	fbController				:FB_STOEBER_AxisController;
	fbMoveManual				:FB_STOEBER_AxisMoveManual;
	fbMoveAuto					:FB_STOEBER_AxisMoveAuto;
	(*fbDriveLink				:FB_STOEBER_DriveLink;*)
	fbForce						:FB_ScalingOffset;
	fbForceCtrl					:FB_ForceController;
	fbCoolingOff				:FB_SignalHandlingDelay;
	
	fbSawingOverride			:FB_Override;
	rtWriteForcePara			:R_TRIG;
	
	fbForceSimple				:FB_ScalingOffset;
	fbForceEL3351				:FB_EL3351;
	fbForceEL3356				:FB_EL3356;

	
END_VAR


IF NOT bEnable								(* Signal FB enable *)
THEN
	bCtrlEnabled := TRUE;
	bReferenced := TRUE;
	bNotMoving := TRUE;
	
	RETURN;
END_IF

A_AxisLink();
A_AxisGetStatus();
A_AxisController();
A_AxisForceCtrl();
A_AxisMoveManual();
A_AxisMoveAuto();
A_AxisTerminalDiag();
A_AxisAlarm();

ACTION A_AxisAlarm:

(* Axis error *)
tonAxisEnabled(
	IN := fbController.bEnable
		AND fbController.bRegulatorOn
		AND NOT fbController.bStatusDelay,
	PT := fbController.tStatusDelay + t#2s
);

bErrorCtrlEnabled := tonAxisEnabled.Q;
(*byErrorPLCOpenController := fbAxisControl.byPLCOpenErrCode;*)
(*bErrorController := fbAxisControl.bError;
bErrorMoveManual := fbMoveManual.bError;
bErrorMoveAuto := fbMoveAuto.bError;*)
END_ACTION

ACTION A_AxisController:

(* Axis controller *)
fbController(
    bEnable := TRUE,
	etMachineMode := etMachineMode,
	etMachineState := etMachineState,
	bNoEStop := bNoEStop,
	bRegulatorOn := bNoEStop
				      AND bPowerSupplyOn
				      AND bSafetyOk
				      AND SEL(bNotMoving, NOT bCtrlInterrupt, TRUE)
				      AND NOT fbMoveManual.bControllerOff
				      AND NOT fbMoveAuto.bControllerOff,
	bReset := bConfirmAlarm,
	bTerminalOK := fbTerminalDiagnosis.bTerminalOK,
	bExeReset := bExeReset,
	bExeSetPos := bExeSetPos,
	lrSetPosition := lrTargetPosition,
	bExeGearIn := bExeGearIn,
	bExeGearOut := bExeGearOut,
	dnRatioNumerator := dnRatioNumerator,
	udnRatioDenominator := udnRatioDenominator,
	lrOverride := SEL(bExtOverrideEn,
					SEL(
						bVeloForceCtrlEn,
						lrOverride,
						fbForceCtrl.lrCVVelo),
					lrOverride*lrExtOverride/100.0)/2,
	bWithAbsoluteEncoder := bWithAbsoluteEncoder,
	bPosLagMonitoringEn := bPosLagMonitoringEn,
	lrPositionBias := lrOriginShiftPos,
	lrSoftLimitMax := lrSoftLimitMax,
	lrSoftLimitMin := lrSoftLimitMin,
	bSignalHWLimitMax:= bSignalHWLimitMax,
	bSignalHWLimitMin := bSignalHWLimitMin,
	lrAcceleration := lrAcceleration,
	lrDeceleration := lrDeceleration,
	lrJerk := lrJerk,
	pDrive := ADR(Drive),
	Axis := Axis,
	MasterAxis := MasterAxis,
	bStatusDelay => bCtrlEnabled,
	lrActPos => lrActPosition,
	lrActAbsPos => lrActAbsPosition,
	lrActVelo => lrActVelocity,
	bNotMoving => bNotMoving,
	bStandStill => bStandStill,
	bReferenced => bReferenced,
	bCoupled => bCoupled,
	lrVeloLimitMax => lrVeloMax,
	lrAccLimitMax => lrAccMax,
	lrDecLimitMax => lrDecMax,
	lrJerkLimitMax => lrJerkMax,
	bHardLimitMaxExceeded => bHardLimitMaxExceeded,
	bHardLimitMinExceeded => bHardLimitMinExceeded,
	bSoftLimitMaxExceeded => bSoftLimitMaxExceeded,
	bSoftLimitMinExceeded => bSoftLimitMinExceeded,

);

bSafetyDriveEnable := fbMoveManual.bSafetyCtrlEnable 
				 	  OR fbMoveAuto.bSafetyCtrlEnable;


(* From Tc2)

(* Sawbow sawing override *)
fbSawingOverride(
	bEnable := bExtOverrideEn
			    AND
			    (etgGr00MachineState = ET_MachineState_eAutoExe
			    OR etgGr00MachineState = ET_MachineState_eAutoSteppingExe)
			    AND
			    (etMachineMode = ET_MachineMode_eAutomatic
			     OR etMachineMode = ET_MachineMode_eCycle
			     OR etMachineMode = ET_MachineMode_eStepping),
	bBypassAccDec := FALSE,
	bSetOverideMax := FALSE,
	rSetOverride := rSetSawingOverride,
	rAcc := rgGr00AdsOverrideAcc,
	rDec := rgGr01AdsOverrideDec
);


IF bExtOverrideEn
     AND
    (etgGr00MachineState = ET_MachineState_eAutoExe
    OR etgGr00MachineState = ET_MachineState_eAutoSteppingExe)
    AND
    (etMachineMode = ET_MachineMode_eAutomatic
     OR etMachineMode = ET_MachineMode_eCycle
     OR etMachineMode = ET_MachineMode_eStepping)
THEN
	rSawingOverride := INT_TO_REAL(nSetSawingOverride)/32767.0 * 100.0;
ELSE
	rSawingOverride := 100.0;
END_IF;

(* Axis controller *)
fbController(
    	bEnable := TRUE,
	etMachineMode := etMachineMode,
	etMachineState := etMachineState,
	bRegulatorOn := bNoEStop
				      AND bPowerSupplyOn
				      AND bSafetyOK
                   		      AND NOT bCtrlInterrupt
				      AND NOT fbMoveManual.bControllerOff
				      AND NOT fbMoveAuto.bControllerOff,
	bReset := bConfirmAlarm,
	bCMDInterrupt := bMoveInterrupt,
	bTerminalOK := fbTerminalDiagnosis.bTerminalOK,
	bExeReset := bExeReset,
  	bExeGearIn := bExeGearIn,
    	bExeGearOut := bExeGearOut,
   	dnRatioNumerator := dnRatioNumerator,
    	udnRatioDenominator := udnRatioDenominator,
	lrOverride := SEL(bExtOverrideEn,
					SEL(
						bVeloForceCtrlEn,
						lrOverride,
						fbForceCtrl.lrCVVelo),
					lrOverride * rSawingOverride / 100),
	lrEngineTorque := SEL(
						bEngineTorqueLimitEn,
						nTorqueLimitMax,
						(lrEngineTorque) / 1),
	bWithAbsoluteEncoder := bWithAbsoluteEncoder,
	bHWSignalLimitMax := bHWSignalLimitMax,
	bHWSignalLimitMin := bHWSignalLimitMin,
	lrSoftLimitMax := lrSoftLimitMax,
	lrSoftLimitMin := lrSoftLimitMin,
	lrAcceleration := lrAcceleration,
	lrDeceleration := lrDeceleration,
	lrJerk := lrJerk,
	tTimeOut := tAdsTimeOut,
	Axis := Axis,
	bStatusDelay => bCtrlEnabled,
	lrActPos => lrActPosition,
	lrActVelo => lrActVelocity,
	bNotMoving => bNotMoving,
	bReferenced => bReferenced,
	bCoupled => bCoupled,
	bHardLimitMaxExceeded => bHardLimitMaxExceeded,
	bHardLimitMinExceeded => bHardLimitMinExceeded,
	bSoftLimitMaxExceeded => bSoftLimitMaxExceeded,
	bSoftLimitMinExceeded => bSoftLimitMinExceeded
);

*)
END_ACTION

ACTION A_AxisForceCtrl:

IF unForceMeasureType = 1			(* Current or voltage force measure *)
THEN
	fbForceCtrl.lrMaxForce := lrForceMaxN; (* [N] *)

	fbForceSimple(
		bEnable := TRUE,
		lrInput := lrForceCurrent,
		lrXLowLimit := lrForceMinmA, (* 16#0000 = 4 [mA] *)
		lrXUpperLimit := lrForceMaxmA, (* 16#7FFF = 20 [mA] *)
		lrYLowLimit := lrForceMinN,  (*[N]*)
		lrYUpperLimit := lrForceMaxN,  (*[N]*)
		usiPrecision := 2,
		lrOffset := rForceOffset,
		lrOutputPV => lrActForce
	);


ELSIF unForceMeasureType = 2			(* EL3351 force measure *)
THEN
	fbForceCtrl.lrMaxForce := lrForceMaxN; (* [N] *)

	fbForceEL3351(
		bEnable := TRUE,
		nTerminalNr := 1,
		stTerminalState := ,
		stBridgeState := ,
		stSupplyState := ,
		dnRefvoltage := ,
		dnDiffvoltage := ,
		rOffset := rForceOffset,
		usiPrecision := 2,
		bDeviceOk => ,
		sDeviceStatus => ,
		rUdiff => ,
		rUref => ,
		lrGrossWeightRV=> ,
		lrGrossWeightPV => lrActForce,
		lrNetWeightRV=> ,
		lrNetWeightPV=> ,
		lrTareWeightRV=> ,
		lrTareWeightPV=>
	);

ELSIF  unForceMeasureType = 3			(* EL3356 force measure *)
THEN

(*
	rtWriteForcePara(
		CLK:= bgGr01ForceActiv5kN
			   XOR bgGr01ForceActiv10kN
	);

	CASE nStepWriteForcePara OF
		0:	(*Idle*)

			fbForceEL3356.bWriteCoePara:= FALSE;
			bWriteForceParaBusy := FALSE;

			IF rtWriteForcePara.Q
			THEN
				nStepWriteForcePara := 10;
				bWriteForceParaBusy := TRUE;
			END_IF
		10: 	(*Start*)

			IF bgGr01ForceActiv5kN
			THEN
				fbForceCtrl.lrMaxForce := 5000, (* [N] *)

				stCoeWrite.bEnableFilter := TRUE;
				stCoeWrite.bEnableUserScale := TRUE;
				stCoeWrite.dwFilterSettings := 0;
				stCoeWrite.rGain := 1.0;
				stCoeWrite.rTara := stgGr01HMI.stHMITOPLC.lrOriginShiftForceX2Right;
				stCoeWrite.rRatedOutput := 0.995000;
				stCoeWrite.rNominalLoad := 5000.0;
				stCoeWrite.rZeroBalance := -0.00028;
				stCoeWrite.rGravityOfEarth := 9.806650;
				stCoeWrite.rScaleFactor := 1.0;
				stCoeWrite.rReferenceLoad	:= 5.0;
				stCoeWrite.bEnableUserScaleIndex8010 := FALSE;
				stCoeWrite.dnUserScaleOffsetIndex8010 := 0;
				stCoeWrite.dnUserScaleGainIndex8010 := 65536;
				stCoeWrite.dwFilterSettingsIndex8010	:= 0;

				fbForceEL3356.bWriteCoePara:= TRUE;

				nStepWriteForcePara := 20;

			ELSIF bgGr01ForceActiv10kN
			THEN
				fbForceCtrl.lrMaxForce := 10000, (* [N] *)

				stCoeWrite.bEnableFilter := TRUE;
				stCoeWrite.bEnableUserScale := TRUE;
				stCoeWrite.dwFilterSettings := 0;
				stCoeWrite.rGain := 1.0;
				stCoeWrite.rTara := stgGr01HMI.stHMITOPLC.lrOriginShiftForceX2Right;
				stCoeWrite.rRatedOutput := 0.9907;
				stCoeWrite.rNominalLoad := 10000.0;
				stCoeWrite.rZeroBalance := 0.00147;
				stCoeWrite.rGravityOfEarth := 9.806650;
				stCoeWrite.rScaleFactor := 1.0;
				stCoeWrite.rReferenceLoad	:= 10.0;
				stCoeWrite.bEnableUserScaleIndex8010 := FALSE;
				stCoeWrite.dnUserScaleOffsetIndex8010 := 0;
				stCoeWrite.dnUserScaleGainIndex8010 := 65536;
				stCoeWrite.dwFilterSettingsIndex8010	:= 0;

				fbForceEL3356.bWriteCoePara:= TRUE;

				nStepWriteForcePara := 20;

			ELSE

				nStepWriteForcePara := 40;
			END_IF

		20: 	(*Wait*)
			IF fbForceEL3356.fbCoe.bCoeBusy
			THEN
				fbForceEL3356.bWriteCoePara:= FALSE;

				nStepWriteForcePara := 30;
			END_IF
	
		30: (*Write*)
			IF NOT fbForceEL3356.fbCoe.bCoeBusy
			THEN
				bWriteForceParaBusy := FALSE;

				IF NOT fbForceEL3356.fbCoe.bCoeError
				THEN
					nStepWriteForcePara := 0;
				ELSE
					nStepWriteForcePara := 40;
				END_IF
			END_IF
		40: (*Error*)
			nStepWriteForcePara := 0;

		ELSE
			nStepWriteForcePara := 0;
	END_CASE

*)

	fbForceCtrl.lrMaxForce := 5000; (* [N] *)

	stCoeWrite.bEnableFilter := TRUE;
	stCoeWrite.bEnableUserScale := TRUE;
	stCoeWrite.dwFilterSettings := 0;
	stCoeWrite.rGain := 1.0;
	stCoeWrite.rTara := (*stgGr01HMI.stHMITOPLC.lrOriginShiftForce*)0.0;
	stCoeWrite.rRatedOutput := 0.995000;
	stCoeWrite.rNominalLoad := 5000.0;
	stCoeWrite.rZeroBalance := -0.00028;
	stCoeWrite.rGravityOfEarth := 9.806650;
	stCoeWrite.rScaleFactor := 1.0;
	stCoeWrite.rReferenceLoad	:= 5.0;
	stCoeWrite.bEnableUserScaleIndex8010 := FALSE;
	stCoeWrite.dnUserScaleOffsetIndex8010 := 0;
	stCoeWrite.dnUserScaleGainIndex8010 := 65536;
	stCoeWrite.dwFilterSettingsIndex8010	:= 0;

	bWriteCoePara := lrCacheWeightTara <> (*stgGr01HMI.stHMITOPLC.lrOriginShiftForce*)0.0;

	fbForceEL3356(
		bEnable := TRUE,
		nTerminalNr := 1,
(*		stTerminalState := stinGr01EL3356A12TerminalState,
		stChannelState := stinGr01EL3356A12ChannelState,*)
		bSetCoeParaToDefault := bSetCoeParaToDefault,
		bReadCoePara := bReadCoePara,
		bWriteCoePara := bWriteCoePara,
		rValue := (*rinGr01ForceRMBValue*)0.0,
		stCoeWrite := stCoeWrite,
		stCoeRead => stCoeRead,
(*		stChannelCtrl => stoutGr01EL3356A8ChannelCtrl,*)
		lrGrossWeightPV =>
	);

	lrActForce := F_LRealRound(fbForceEL3356.lrGrossWeightPV - rForceOffset, 2);

	lrCacheWeightTara := (*stgGr01HMI.stHMITOPLC.lrOriginShiftForce*)0.0;

ELSE							(* Directly force measure *)

	lrActForce := lrForceCurrent;
	fbForceCtrl.lrMaxForce := lrForceMaxN; (* [N] *)

END_IF

fbForceCtrl(
	bEnable := bNoEStop
			    AND bPowerSupplyOn
			    AND bSafetyOK
			    AND bCtrlEnabled,
	bControllerOn := bVeloForceCtrlEn,
	lrVeloKp := lrVeloForceCtrlKp,
	lrVeloTi := lrVeloForceCtrlTi,
	lrCtrlVeloFilter := lrVeloForcePreCtrlVelo,
	lrPVForce := lrActForce, (* [N] *)
	lrSPForce := lrTargetForce, (* [N] *)
	lrVeloMax := lrVeloForceCtrlMax,
	lrVeloMin := lrVeloForceCtrlMin,
	lrTaskCycle := lrgActCycleTime
);
END_ACTION

ACTION A_AxisGetStatus:

(* Get axis status *)
Axis.ReadStatus();
END_ACTION

ACTION A_AxisLink:

(* Get terminal status *)
sAdsAddr := F_CreateAmsNetId(Drive.stTerminalState.stAdsAddr.netId);
unSlaveAddr := Drive.stTerminalState.stAdsAddr.port;
Axis.DriveAddress.NetID := F_CreateAmsNetId(Drive.stTerminalState.stAdsAddr.netId);
Axis.DriveAddress.SlaveAddress := Drive.stTerminalState.stAdsAddr.port;

(* Set drive parameter *)
Drive.stPlcToStoeber.snA541ModesOfOperation := snModesOfOperation;

(*Drive.PlcToStoeber.nA558TargetTorque := SEL(bEngineTorqueLimitEn,
				    nTorqueLimitMax,
				    LREAL_TO_INT(lrEngineTorque / 1.0))*)
END_ACTION

ACTION A_AxisMoveAuto:

(* Move axis auto *)
rtMachineStandstill(CLK := bMachineStandstill);

lrVeloLimitMin := SEL(bVelocityLimitEn, -1 * lrVeloMax, lrVelocityMin);
lrVeloLimitMax := SEL(bVelocityLimitEn, lrVeloMax, lrVelocityMax);;

fbMoveAuto(
	bEnable := bNoEStop
               		    AND bPowerSupplyOn
               		    AND bSafetyOK,
    	bCtrlEnabled := bCtrlEnabled
                    		   AND bMoveRelease,
	etMachineMode := etMachineMode,
	etMachineState := etMachineState,
	bReset := bConfirmAlarm,
	bExeHome := bExeHome,
	bExeMoveAbs := bExeMoveAbs,
	bExeMoveRel := bExeMoveRel,
	bExeMoveAdd := bExeMoveAdd,
	bExeMoveSuper := bExeMoveSuper,
	bExeMoveVelo := bExeMoveVelo,
	bExeStop := bExeStop
			      OR rtMachineStandstill.Q,
	lrPosition := lrTargetPosition,
	lrVelocity := LIMIT(lrVeloLimitMin, lrAutoVelocity, lrVeloLimitMax),
	lrAcceleration := lrAcceleration,
	lrDeceleration := lrDeceleration,
	lrJerk := lrJerk,
	lrOriginShiftPos := lrOriginShiftPos,
	bSignalReference := bSignalReference,
	tControllerOff := tControllerOff,
	bHomeCompleted := bHomeCompleted,
	Axis := Axis,
	MasterAxis 				:= GVL_Gr00Interface.iAxisDummy,
 );
END_ACTION

ACTION A_AxisMoveManual:

(* Move axis manual *)
fbMoveManual(
	bEnable := bNoEStop
               AND bPowerSupplyOn
               AND bSafetyOK,
	bOccupied := bOccupied,
	bSafetyCtrlEnabled := bSafetyDriveEnabled,
	bCtrlEnabled := bCtrlEnabled
				    AND bMoveRelease,
	etMachineMode := etMachineMode,
	etMachineState := etMachineState,
	bReset := bConfirmAlarm,
	bMovePlus := bTipPlus,
	bMoveMinus := bTipMinus,
	lrTipDistance := lrTipDistance,
	bLimitMax := bHardLimitMaxExceeded
			     OR bSoftLimitMaxExceeded,
	bLimitMin := bHardLimitMinExceeded
			     OR bSoftLimitMinExceeded,
	bPlusRelease := bPlusRelease,
	bMinusRelease := bMinusRelease 
					 AND NOT bErrorForceOverflow,
	lrVelocity := SEL(NOT bReferenced, lrManualVelocity, lrNoRefVelocity),
	lrAcceleration := lrAcceleration,
	lrDeceleration := lrDeceleration,
	lrJerk := lrJerk,
	tControllerOff := tControllerOff,
	pDrive := ADR(Drive),
	bHomeCompleted := bHomeCompleted,
	Axis := Axis,
	MasterAxis := MasterAxis
);

(* From Tc2)
(* Move axis manual *)
fbMoveManual(
	bEnable := bNoEStop
               		    AND bPowerSupplyOn
               		    AND bSafetyOK,
	bCtrlEnabled := bCtrlEnabled
                			    AND bMoveRelease,
	etMachineMode := etMachineMode,
	etMachineState := etMachineState,
	bReset := bConfirmAlarm,
	bMovePlus := bTipPlus,
	bMoveMinus := bTipMinus,
	lrTipDistance := lrTipDistance,
	bLimitMax := bHardLimitMaxExceeded
			       OR bSoftLimitMaxExceeded ,
	bLimitMin := bHardLimitMinExceeded
			      OR bSoftLimitMinExceeded,
	bPlusRelease := bPlusRelease,
	bMinusRelease := bMinusRelease,
	lrVelocity := SEL(NOT bReferenced, lrManualVelocity, lrVelocityNoRef),
	lrAcceleration := lrAcceleration,
	lrDeceleration := lrDeceleration,
	lrJerk := lrJerk,
	tControllerOff := tControllerOff,
	bHomeCompleted := bHomeCompleted,
	Axis := Axis
);

bSafetyLock := fbMoveManual.bMovePlus
                		OR fbMoveManual.bMoveMinus;
						
*)
END_ACTION

ACTION A_AxisTerminalDiag:

(*Axis terminal diagnosis *)
fbTerminalDiagnosis(
	stTerminalState := Drive.stTerminalState,
	sTerminalStatus => sTerminalStatus
);

bErrorTerminal := NOT fbTerminalDiagnosis.bTerminalOK;
END_ACTION

END_FUNCTION_BLOCK

// ---- POUs/Tc2 Objects/Diagnostic/Terminal/FB_TerminalDiagnosis.TcPOU
FUNCTION_BLOCK FB_TerminalDiagnosis
VAR_INPUT
	stTerminalState				:ST_TerminalState;
END_VAR
VAR_OUTPUT
	bTerminalOK					:BOOL;
	sTerminalStatus				:STRING;
END_VAR
VAR

	sStateStatusAll				:STRING(255);
	sState						:STRING;
	sWorkingState				:STRING;
	tonTerminalNOK				:TON;
END_VAR
VAR CONSTANT
	tTerminalNOKDelay				:TIME := t#2s;
END_VAR

(*This Function returns the State of the Device. Either one of the States INIT, PREOP, OP, BOOTSTRAP or SAFE-OP is returned. stState is given the Value of the Function. *)
sState:= F_StateReturn(state:= stTerminalState.unInfoState);

(*All other Errors that can occur concerning the State of the Device*)
(*Because theoratically all the other errors could occur all together, CONCAT is done to show them all in one view box.*)
IF stTerminalState.unInfoState.4
THEN
	sStateStatusAll:= 'Slave signals error. ';
ELSE
	sStateStatusAll:= '';
END_IF

IF stTerminalState.unInfoState.5
THEN
	sStateStatusAll:= CONCAT( sStateStatusAll, 'Invalid vendorID. ');
ELSE
	sStateStatusAll:= CONCAT( sStateStatusAll, '');
END_IF

IF stTerminalState.unInfoState.6
THEN
	sStateStatusAll:= CONCAT( sStateStatusAll, 'Initialization error occurred. ');
ELSE
	sStateStatusAll:= CONCAT( sStateStatusAll, '');
END_IF

IF stTerminalState.unInfoState.7
THEN
	sStateStatusAll:= CONCAT( sStateStatusAll, 'Slave disabled. ');
ELSE
	sStateStatusAll:= CONCAT( sStateStatusAll, '');
END_IF

IF stTerminalState.unInfoState.8
THEN
	sStateStatusAll:= CONCAT( sStateStatusAll, 'Slave not present. ');
ELSE
	sStateStatusAll:= CONCAT( sStateStatusAll, '');
END_IF

IF stTerminalState.unInfoState.9
THEN
	sStateStatusAll:= CONCAT( sStateStatusAll, 'Slave signals link error. ');
ELSE
	sStateStatusAll:= CONCAT( sStateStatusAll, '');
END_IF

IF stTerminalState.unInfoState.10
THEN
	sStateStatusAll:= CONCAT( sStateStatusAll, 'Slave signals missing link. ');
ELSE
	sStateStatusAll:= CONCAT( sStateStatusAll, '');
END_IF

IF stTerminalState.unInfoState.11
THEN
	sStateStatusAll:= CONCAT( sStateStatusAll, 'Slave signals unexpected link. ');
ELSE
	sStateStatusAll:= CONCAT( sStateStatusAll, '');
END_IF

IF stTerminalState.unInfoState.12
THEN
	sStateStatusAll:= CONCAT( sStateStatusAll,  'Communication port A. ');
ELSE
	sStateStatusAll:= CONCAT( sStateStatusAll, '');
END_IF

IF stTerminalState.unInfoState.13
THEN
	sStateStatusAll:= CONCAT( sStateStatusAll, 'Communication port B. ');
ELSE
	sStateStatusAll:= CONCAT( sStateStatusAll, '');
END_IF

IF stTerminalState.unInfoState.14
THEN
	sStateStatusAll:= CONCAT( sStateStatusAll, 'Communication port C. ');
ELSE
	sStateStatusAll:= CONCAT( sStateStatusAll, '');
END_IF

IF stTerminalState.unInfoState.15
THEN
	sStateStatusAll:= CONCAT( sStateStatusAll,  'Communication port D. ');
ELSE
	sStateStatusAll:= CONCAT( sStateStatusAll, '');
END_IF

(*If none of the other errors occur, the text of the view box is 'None'.*)
IF sStateStatusAll= ''
THEN
	sStateStatusAll:= 'No error';
END_IF

(*The colour and text of the view box WcState is adjusted.*)
IF stTerminalState.bWcState = 0
THEN
	sWorkingState:= 'Working State OK ';
ELSE
	sWorkingState:= 'Working State NOT OK ';
END_IF

(*General Status Information*)
bTerminalOK:= TRUE;
sTerminalStatus:= 'Terminal OK ';

IF stTerminalState.bWcState <> 0
     OR sStateStatusAll <> 'No error'
THEN
	tonTerminalNOK(IN := TRUE, PT := tTerminalNOKDelay);
	IF tonTerminalNOK.Q
	THEN
		bTerminalOK:= FALSE;
		sTerminalStatus:= 'Terminal Error ';
	ELSE
		sTerminalStatus:= 'Waiting for status.';
	END_IF
END_IF

END_FUNCTION_BLOCK

// ---- POUs/Tc2 Objects/Diagnostic/Terminal/F_StateReturn.TcPOU
FUNCTION F_StateReturn : STRING
VAR_INPUT
	state: UINT;
END_VAR
VAR
END_VAR

(*This Function returns the State of the Device. Either one of the States INIT, PREOP, OP, BOOTSTRAP or SAFE-OP is returned.
FB_Diagnosis.stState is given the Value of this Function. *)

IF state.0 AND NOT state.1 THEN
	F_StateReturn:= 'Slave in INIT state';
END_IF
IF state.1 AND NOT state.0 THEN
	F_StateReturn:= 'Slave in PREOP state';
END_IF
IF state.0 AND state.1 THEN
	F_StateReturn:= 'Slave in BOOTSTRAP state';
END_IF
IF state.2 THEN
	F_StateReturn:= 'Slave in SAFEOP state';
END_IF
IF state.3 THEN
	F_StateReturn:= 'Slave in OP state';
END_IF

END_FUNCTION

// ---- POUs/Tc2 Objects/Mathematical/Scaling/FB_ScalingOffset.TcPOU
FUNCTION_BLOCK FB_ScalingOffset
(*

The function block used to scaling input signal.

Constructor: 		Patryk Panylo
Company:		E. Riexinger GmbH
Date:			04.08.2015
Version:			1.00

Date:			Revision:		Who:				Comment
dd.mm.yyyy		x.xx			Initials			comment

*)
VAR_INPUT
	(* Input variables / Eingang Variablen *)
	bEnable							:BOOL;						(* Function block enable *)
	lrInput							:LREAL;						(* Input scaling proces value *)
	lrXLowLimit						:LREAL;						(* Upper limit of X range *)
	lrXUpperLimit						:LREAL; 						(*Upper limit of X range  *)
	lrYLowLimit						:LREAL; 						(* Low limit of Y range  *)
	lrYUpperLimit						:LREAL; 						(* Upper limit of Y range  *)
	usiPrecision						:USINT := 2; 					(* The number of digits after the decimal point depends on the requested precision *)
	lrOffset							:LREAL;						(* Offset of output *)
END_VAR
VAR_OUTPUT
	(* Output variables / Ausgang Variablen *)
	lrOutputRV						:LREAL;						(* Raw Value *)
	lrOutputPV						:LREAL;						(* Judgment Value  *)
END_VAR
VAR
	(* Instances / Instanzen *)
	fbScaling						:FB_Scaling;

	(* Enumerator  *)

	(* General flags / Allgemeine Variablen *)

END_VAR
VAR CONSTANT

END_VAR

IF NOT bEnable THEN
	fbScaling(
		bEnable := FALSE,
	);

	lrOutputRV := 0.0;					(* Raw Value *)
	lrOutputPV := 0.0;					(* Judgment Value *)
	RETURN;
END_IF

(* Scaling *)

fbScaling(
	bEnable := TRUE,
	lrInput := lrInput,
	lrXLowLimit := lrXLowLimit,
	lrXUpperLimit := lrXUpperLimit,
	lrYLowLimit := lrYLowLimit,
	lrYUpperLimit := lrYUpperLimit,
	usiPrecision := usiPrecision
);

lrOutputRV := fbScaling.lrOutputRV + lrOffset;
lrOutputPV := fbScaling.lrOutputPV + lrOffset;

END_FUNCTION_BLOCK

// ---- POUs/Tc2 Objects/Mathematical/Scaling/FB_Scaling.TcPOU
FUNCTION_BLOCK FB_Scaling
(*

The function block used to scaling input signal.

Constructor: 		Patryk Panylo
Company:		E. Riexinger GmbH
Date:			04.08.2015
Version:			1.00

Date:			Revision:		Who:				Comment
dd.mm.yyyy		x.xx			Initials			comment

*)
VAR_INPUT
	(* Input variables / Eingang Variablen *)
	bEnable							:BOOL;						(* Function block enable *)
	lrInput							:LREAL;						(* Input scaling proces value *)
	lrXLowLimit						:LREAL;						(* Upper limit of X range *)
	lrXUpperLimit						:LREAL; 						(*Upper limit of X range  *)
	lrYLowLimit						:LREAL; 						(* Low limit of Y range  *)
	lrYUpperLimit						:LREAL; 						(* Upper limit of Y range  *)
	usiPrecision						:USINT := 2; 					(* The number of digits after the decimal point depends on the requested precision *)
END_VAR
VAR_OUTPUT
	(* Output variables / Ausgang Variablen *)
	lrOutputRV						:LREAL;						(* Raw Value *)
	lrOutputPV						:LREAL;						(* Judgment Value  *)
	bLowLevel						:BOOL;						(* Low level detected *)
	bGoLevel						:BOOL;						(* Go level detected *)
	bHighLevel						:BOOL;						(* High level detected *)
END_VAR
VAR
	(* Instances / Instanzen *)

	(* Enumerator  *)

	(* General flags / Allgemeine Variablen *)
	lra								:LREAL;
	lrb								:LREAL;
END_VAR
VAR CONSTANT

END_VAR

IF NOT bEnable THEN
	lrOutputRV := 0.0;					(* Raw Value *)
	lrOutputPV := 0.0;					(* Judgment Value *)
	bLowLevel := FALSE;				(* Low level detected *)
	bGoLevel := FALSE;					(* Go level detected *)
	bHighLevel := FALSE;				(* High level detected *)
	RETURN;
END_IF

(* Scaling *)
IF lrInput > lrXUpperLimit															(* Check upper limit of X range *)
THEN
	lrOutputRV := lrYUpperLimit;
	bLowLevel := FALSE;
	bHighLevel := TRUE;
	bGoLevel := FALSE;
ELSIF lrInput <= lrXLowLimit														(* Check low limit of X range *)
THEN
	lrOutputRV := lrYLowLimit;
	bLowLevel := TRUE;
	bHighLevel := FALSE;
	bGoLevel := FALSE;
ELSE
	IF (((lrXUpperLimit - lrXLowLimit) < 0.01)											(* Check X range *)
	    AND ((lrXUpperLimit - lrXLowLimit) > -0.01))
	THEN
		lrOutputRV := lrYLowLimit;
		bLowLevel := TRUE;
		bHighLevel := FALSE;
		bGoLevel := FALSE;
	ELSE
		lra := (lrYUpperLimit - lrYLowLimit) / (lrXUpperLimit - lrXLowLimit);					(* Slope of a straight line, drawed by the range positions *)
		lrb := lrYUpperLimit - lra * lrXUpperLimit;
		lrOutputRV := lra * lrInput + lrb;
		bLowLevel := FALSE;
		bHighLevel := FALSE;
		bGoLevel := TRUE;
	END_IF;
END_IF

lrOutputPV := F_LRealRound(lrOutputRV, usiPrecision);

END_FUNCTION_BLOCK

// ---- POUs/Tc2 Objects/Mathematical/F_LRealRound.TcPOU
FUNCTION F_LRealRound : LREAL
(*

The function used to round lreal value.

Constructor: 		Patryk Panylo
Company:		E. Riexinger GmbH
Date:			04.08.2015
Version:			1.00

Date:			Revision:		Who:				Comment
dd.mm.yyyy		x.xx			Initials			comment

*)
VAR_INPUT
	(* Input variables / Eingang Variablen *)
	lrReal							:LREAL; 						(*  Input variable *)
	usiPrecision						:USINT := 2; 					(* The number of digits after the decimal point depends on the requested precision *)
END_VAR
VAR
	(* Variables *)
	lrFraction							:LREAL;
END_VAR

(* Round real value with precision *)
lrFraction := FRAC(ABS(lrReal)) * EXPT(10, usiPrecision + 1); 							(* The fraction of the value *)

IF LMOD(lrFraction, 10) < 5
THEN
	lrFraction := lrFraction - LMOD(lrFraction, 10) ;										(* Round down *)
ELSE
	lrFraction := lrFraction + (10 - LMOD(lrFraction, 10));									(* Round up and check the integral increment *)
END_IF;

IF lrReal  < 0																		(* Check the digit of the value *)
THEN
	F_LRealRound	 := LTRUNC(lrReal) - (lrFraction / EXPT(10, usiPrecision + 1));
ELSE
	F_LRealRound	 := LTRUNC(lrReal) + (lrFraction / EXPT(10, usiPrecision + 1));
END_IF

END_FUNCTION

// ---- POUs/Tc2 Objects/Automation/Force/FB_ForceController.TcPOU
FUNCTION_BLOCK FB_ForceController
(*

The function block used to 

Constructor: 		Patryk Panylo
Company:		E. Riexinger GmbH
Date:			17.02.2016
Version:			1.00

Date:			Revision:		Who:				Comment

*)
VAR_INPUT
	(* Input variables / Eingang Variablen *)
	bEnable					:BOOL;					(* Signal FB enable *)
	bControllerOn				:BOOL;					(* Controler on *)
	lrVeloKp					:LREAL := 0.1;				(* Kp Proportionalfaktor, deltaF x Kp -> v *)
	lrVeloTi					:LREAL := 10000;			(* Ti Integrationsfaktor*)
	lrCtrlVeloFilter				:LREAL := 0.01;			(* Control velocity filter =  0..1 *)
	lrPVForce				:LREAL;					(* Process variable of force *)
	lrSPForce				:LREAL;					(* Set point of force *)
	lrMaxForce				:LREAL;					(* Maximum force *)
	lrDeltaMax				:LREAL := 0.01;
	lrVeloMax				:LREAL := 10.0;			(* Maximum velocity [%] *)
	lrVeloMin				:LREAL := 0.0;				(* Minimum velocity [%] *)
	lrTaskCycle				:LREAL;					(* Task cycle *)
END_VAR
VAR_OUTPUT
	(* Output variables / Ausgang Variablen *)
	lrCVVelo					:LREAL;					(* Controller value of velocity [%] *)
END_VAR
VAR_IN_OUT
	(* Input Output variables / Ausgang Variablen *)

END_VAR
VAR
	(* Enummerations *)

	(* Variables *)

	(* References *)

	(* Interfaces *)

	(* Instances *)
	fbActForceFilter				:FB_ValueFilter;					(* Actual position filter *)
	fbCtrlPID						:FB_CtrlPID;

END_VAR
VAR CONSTANT

END_VAR


IF NOT bEnable
THEN
	lrCVVelo := 100;
	RETURN;
END_IF

(* Current force value filtering *)
fbActForceFilter(
	bEnable := TRUE,
	lrInSignal := lrPVForce,
	lrDeltaMax := lrDeltaMax,
);

IF bControllerOn
     AND fbActForceFilter.lrOutSignal < lrMaxForce
THEN

	fbCtrlPID(
		bEnable := TRUE,
		lrSetPoint := lrSPForce,
		lrProcessVariable := fbActForceFilter.lrOutSignal,
		lrDeadZone := 1.0,
		lrSignalOffset := 0.0,
		lrKp := lrVeloKp,
		lrTi := lrVeloTi,
		lrTd := 0.0,
		lrTaskCycle := lrTaskCycle,
		bManual := ,
		lrManualSignal:= ,
		lrLimitMin := lrVeloMin,
		lrLimitMax := lrVeloMax,
		lrProcessErr => ,
		bLimitMin => ,
		bLimitMax => );


	(*Reg_Rueck := Reg_Filt*Reg_Rueck + (1-Reg_Filt)*Reg_Verst*Drehzahl*Y_Vmax;*)
	(*lrCVVelo := MAX(0.0, (fbCtrlPID.lrCtrlVariable * (1.0 - lrPreCtrlVelo)) + (fbActForceFilter.lrOutSignal * lrPreCtrlVelo)); (* where lrPreCtrlVelo := 0.01 *)*)
	(*lrCVVelo := MAX(0.0, (fbCtrlPID.lrCtrlVariable * (1.0 - lrCtrlVeloFilter)) + (lrCVVelo * lrCtrlVeloFilter));				       (* where lrPreCtrlVelo := 0.99 *)*)
	lrCVVelo := MAX(0.0, (fbCtrlPID.lrCtrlVariable * lrCtrlVeloFilter) + (lrCVVelo * (1.0 - lrCtrlVeloFilter)));				       (* where lrPreCtrlVelo := 0.99 *)

ELSE
	lrCVVelo := 0.0;
END_IF

END_FUNCTION_BLOCK

// ---- POUs/Tc2 Objects/Engineering/Filter/FB_ValueFilter.TcPOU
FUNCTION_BLOCK FB_ValueFilter
(*

Function block for filtering current input-value.

Sample Time
Constructor: 		Patryk Panylo
Company:		E. Riexinger GmbH
Date:			16.07.2014
Version:			1.00

Date:			Revision:		Who:				Comment
dd.mm.yyyy		x.xx			Initials			comment

*)
VAR_INPUT
	(* Enummerations *)

	(* Variables *)
	bEnable								:BOOL := TRUE;					(* Enable FB *)

	lrInSignal								:LREAL;							(* Input signal *)
	lrDeltaMax							:LREAL := 100;					(* Maximum difference between two input values *)

	(* References *)

	(* Interfaces *)

	(* Instances *)

END_VAR
VAR_OUTPUT
	(* Enummerations *)
	
	(* Variables *)
	lrOutSignal							:LREAL;							(* Output signal *)

	(* References *)

	(* Interfaces *)

	(* Instances *)
END_VAR
VAR
	(* Enummerations *)
	
	(* Variables *)
	bFirstTime							:BOOL;							(* First cycle *)

	lrCacheInSignal						:LREAL;							(* Copy of input signal *)
	dnOverLimitCounter					:DINT;							(* Counter of over limit *)

	lrLastSignal							:LREAL;							(* Last signal in time N *)
	lrSignalN_1							:LREAL;							(* Signal in time N - 1 *)
	lrSignalN_2							:LREAL;							(* Signal in time N - 2 *)
	lrSignalN_3							:LREAL;							(* Signal in time N - 3 *)

	(* References *)

	(* Interfaces *)

	(* Instances *)




END_VAR

IF NOT bEnable
THEN
	lrOutSignal := lrInSignal;

	bFirstTime := FALSE;
	RETURN;
END_IF

IF NOT bFirstTime
THEN
	lrSignalN_3 := lrInSignal;
	lrSignalN_2 := lrInSignal;
	lrSignalN_1 := lrInSignal;
	lrLastSignal := lrInSignal;

	bFirstTime := TRUE;
END_IF

lrSignalN_3 := lrSignalN_2;
lrSignalN_2 := lrSignalN_1;
lrSignalN_1 := lrLastSignal;

lrCacheInSignal := lrInSignal;

IF ABS( lrCacheInSignal - lrSignalN_1 ) <= lrDeltaMax
THEN
	lrLastSignal := lrCacheInSignal;
	dnOverLimitCounter := 0;

ELSE
	dnOverLimitCounter := dnOverLimitCounter + 1;

	IF dnOverLimitCounter <= 3
	THEN
		lrLastSignal	:= lrSignalN_1 + ((lrSignalN_1 - lrSignalN_2) + (lrSignalN_2 - lrSignalN_3)) / 2.0;

	ELSIF dnOverLimitCounter = 4
	THEN
		lrLastSignal := lrSignalN_1 + (lrCacheInSignal - lrSignalN_1) / 2.0;

	ELSE
		lrLastSignal := lrCacheInSignal;
	END_IF

END_IF

lrOutSignal := lrLastSignal;

END_FUNCTION_BLOCK

// ---- POUs/Machine/Group_0100 - Production/Gr01Control/Gr01Units/FB_Gr01Angle.TcPOU
FUNCTION_BLOCK FB_Gr01Angle
(*

The function block used to control axis .

Constructor: 		Patryk Panylo
Company:		E. Riexinger GmbH
Date:			28.04.2015
Version:			1.00

Date:			Revision:		Who:				Comment
dd.mm.yyyy		x.xx			Initials			comment

*)
VAR_INPUT
	(* Input variables / Eingang Variablen *)
	(* --- Axis / Achse --- *)
	bEnable						:BOOL;						(* Axis present *)
	bOccupied					:BOOL;						(* Axis is occupied *)

	(* --- Machine state / Maschinenzustand --- *)
	etMachineMode				:ET_MachineMode;			(* Machine mode *)
	etMachineState				:ET_MachineState;			(* Machine state *)
	bMachineStandstill			:BOOL;						(* Machine standstill *)

	(* --- Safety & releases / Sicherheit & Freigaben --- *)
	bNoEStop					:BOOL;						(* No ermergency Stop / Keine Notaus *)
	bPowerSupplyOn				:BOOL;						(* Power supply on / Leitung eingeschaltet *)
	bSafetyOK					:BOOL;						(* Safety ok / Sicherheit i.o *)
	bSafetyDriveEnabled			:BOOL;						(* Safety drive enable *)
	bCtrlInterrupt				:BOOL;						(* Control interrupt *)
	bMoveRelease				:BOOL;						(* Move release *)
	bMoveInterrupt				:BOOL;						(* Move Interrupt *)
	bPlusRelease				:BOOL;						(* Plus move release *)
	bMinusRelease				:BOOL;						(* Minus move release *)

	(* --- Limits / Endlagen --- *)
	bHWSignalLimitMax			:BOOL;						(* Signal position limit switch maximum *)
	bHWSignalLimitMin			:BOOL;						(* Signal position limit switch minimum *)
	lrSoftLimitMax				:LREAL;						(* Position limit switch maximum *)
	lrSoftLimitMin				:LREAL;						(* Position limit switch minimum *)

	(* --- Commands / Befehle --- *)
	bExeReset					:BOOL;						(* Execute auto reset *)
	bExeHome					:BOOL;						(* Execute home *)
	bExeMoveAbs					:BOOL;						(* Execute move absolut *)
	bExeMoveVelo				:BOOL;						(* Execute move velo *)
	bExeGearIn					:BOOL;						(* Execute gear in *)
	bExeGearOut					:BOOL;						(* Execute gear out *)
	bExeStop					:BOOL;						(* Execute move stop *)
	bConfirmAlarm				:BOOL;						(* Confirm alarm *)

	(* --- Manual mode / Handbetrieb --- *)
	bTipPlus					:BOOL;						(* Manual tip in plus direction *)
	bTipMinus					:BOOL;						(* Manual tip in minus direction *)
	lrManualVelocity			:LREAL;						(* Value of velocity in manual motion [mm/s] *)

	(* --- Motion parameters / Bewegungsparameter --- *)
	lrTargetPosition			:LREAL;						(* Absolute target position *)
	lrAutoVelocity				:LREAL;						(* Value of velocity in auto motion [mm/s] *)
	lrVelocityNoRef				:LREAL;						(* Velocity if has no reference [mm/s] *)
	bVelocityLimitEn			:BOOL;						(* Enable velocity limit *)
	lrVelocityMin				:LREAL;						(* Velocity minimum [%] *)
	lrVelocityMax				:LREAL;						(* Velocity maximum [%] *)
	lrAcceleration				:LREAL;						(* Value of the acceleration (always positive) *)
	lrDeceleration				:LREAL;						(* Value of deceleration (always positive) *)
	lrJerk						:LREAL;						(* Value of jerk (always positive) *)

	(* --- Override --- *)
	lrOverride					:LREAL;						(* Override *)
	bExtOverrideEn				:BOOL;						(* External override enable *)
	lrExtOverride				:LREAL;						(* External override *)

	(* --- Gearing / Getriebe --- *)
	dnRatioNumerator			:DINT;						(* Gear ratio numerator. Alternatively, the gear ratio can be specified in the numerator as a floating comma value, if the denominator is 1. *)
	udnRatioDenominator			:UDINT;						(* Gear ratio denominator *)

	(* --- Drive / Antrieb --- *)
	snModesOfOperation			:SINT;						(* Modes of drive operation *)
	bEngineTorqueLimitEn		:BOOL;						(* Enable engine torque limit *)
	lrEngineTorque				:LREAL;						(* Engine torque [%] *)
	bPosLagMonitoringEn			:BOOL;						(* Enable position lag monitoring *)
	tControllerOff				:TIME := T#60S;				(* Time to switch controller off *)

	(* --- Scaling & encoder / Skalierung & Geber --- *)
	lrScalingNum				:LREAL := 1.0;				(* Effective distance per rev. Numerator [technical units] *)
	udnScalingDenom				:UDINT := 1;				(* Effective distance per rev. Denominator [INC] *)
	bWithAbsoluteEncoder		:BOOL;						(* Encoder is an absolute one / Absolutwertgeber *)
	udnIncEnc					:UDINT;						(* Value of encoder increment *)
	lrOriginShift				:LREAL;						(* Origin shift position *)

	(* --- System --- *)
	lrTaskCycle					:LREAL := 0.002;			(* Cycle time of the task [sec], 0.002[s] => 2ms *)
	tAdsTimeOut					:TIME := T#2S;				(* Timout for ads commands *)
END_VAR
VAR_OUTPUT
	(* Output variables / Ausgang Variablen *)
	(* --- Status --- *)
	bCtrlEnabled				:BOOL;						(* Controller enabled *)
	bNotMoving					:BOOL;						(* Axis not moving *)
	bStandStill					:BOOL;						(* Added by Dustin for 633_Hilton) Axis stands stil*)
	bReferenced					:BOOL;						(* Axis referenced *)
	bCoupled					:BOOL;						(* Axis coupled *)

	(* --- Actual values / Istwerte --- *)
	lrActPosition				:LREAL;						(* Actual position [mm] *)
	lrActAbsPosition			:LREAL;						(* Actual absolut position [mm] *)
	lrActVelocity				:LREAL;						(* Actual velocity [mm/s] *)
	lrVeloMax					:LREAL;						(* Velocity limit maximum *)

	(* --- Limits / Endlagen --- *)
	bHardLimitMaxExceeded		:BOOL;						(* Position limit switch maximum is exceeded *)
	bHardLimitMinExceeded		:BOOL;						(* Position limit switch minimum is exceeded *)
	bSoftLimitMaxExceeded		:BOOL;						(* Position limit switch maximum is exceeded *)
	bSoftLimitMinExceeded		:BOOL;						(* Position limit switch minimum is exceeded *)

	(* --- Safety / Sicherheit --- *)
	bSafetyLock					:BOOL;						(* Safety lock*)
	bSafetyDriveEnable			:BOOL;						(* Safety drive enable *)

	(* --- Errors / Fehler --- *)
	bErrorTerminal				:BOOL;						(* Error Axis terminal *)
	bErrorCtrlEnabled			:BOOL;						(* Error Axis controller enabled *)
	
END_VAR
VAR_IN_OUT	
	(* Input Output variables / Ausgang Variablen *)
	bHomeCompleted				:BOOL;						(* Home completed *)
	Drive						:ST_STOEBERSI6SC6CIA402_REF;
	Axis						:AXIS_REF;
	MasterAxis					:AXIS_REF;
END_VAR
VAR
	(* Enummerations *)

	(* Variables *)
	sAdsAddr					:STRING(23);					(* AmsNetId of the EtherCAT master device.*)
	unSlaveAddr					:UINT;							(* Address of the slave device.*)

	nTorqueLimitMax				:INT := 100;					(* The torque limit (absolute value). Value range in %: -200 ... 200 ... 200 *)

	lrVeloLimitMax				:LREAL;
	lrVeloLimitMin				:LREAL;

	sTerminalStatus				:STRING;

	(* References *)

	(* Interfaces *)

	(* Instances *)
	fbTerminalDiagnosis			:FB_TerminalDiagnosis;
	rtMachineStandstill			:R_TRIG;
	tonAxisEnabled				:TON;

	fbController				:FB_STOEBER_AxisController;
	fbMoveManual				:FB_STOEBER_AxisMoveManual;
	fbMoveAuto					:FB_STOEBER_AxisMoveAuto;
	(*fbDriveLink				:FB_STOEBER_DriveLink;*)
	fbForce						:FB_ScalingOffset;
	fbForceCtrl					:FB_ForceController;
	fbCoolingOff				:FB_SignalHandlingDelay;
END_VAR


IF NOT bEnable								(* Signal FB enable *)
THEN

	RETURN;
END_IF

(* Old Axis Ref from Tc2) 
(* ControllerConfig *)
stControllerConfig.lrKp := 0.018;						(* Tuning parameter, proportional gain *)
stControllerConfig.lrTi := 0.0;							(* Tuning parameter, time of integral *)
stControllerConfig.lrTd := 0.0;						(* Tuning parameter, time of differential *)
stControllerConfig.lrPreCtrlVelo := 0.01; 				(* Feedforward velocity precontrol wieghting =  0..1 *)
stControllerConfig.lrVeloKpFilter := 1.0;				(* Velocity filter - proportional gain *)
stControllerConfig.tVeloT1Filter := t#100ms;			(* Velocity filter - time constant *)
stControllerConfig.tDeadTime  := t#100ms;				(* Dead time *)
stControllerConfig.lrDeltaMax := 10.0;					(* Maximum difference between two actual position values filtered [inc] *)
stControllerConfig.lrVeloMin := -7.8; 					(* Velocity limit minimum [deg / sec] *)
stControllerConfig.lrVeloMax  := 7.8; 					(* Velocity limit maximum [deg / sec] *)
stControllerConfig.lrDeadZone := 10.0;					(* Dead zone *)

(* Encoder configuration *)
stEncoderConfig.dwModuloValue := 8192; 			(* Maximum encoder modulo value e.g 1048576 [inc] *)
stEncoderConfig.etScalingMethod := ET_ScalingMethod_eSMLinear;

(* Interface *)
stAxis.stScaling.dwModuloValue := 8192; 		(* Maximum encoder modulo value 4294967295 dword *)
stAxis.stAxisCtrl.bEnable := Axis.stPlcToNc.stBaseDevice.bEnable;
stAxis.stAxisStates.bOperational := Axis.stNcToPlc.stBaseDevice.bEnabled;
stAxis.stScaling.etScalingMethod := ET_ScalingMethod_eSMLinear;
stAxis.stScaling.lrTaskCycle := lrTaskCycle;
stAxis.stScaling.udnScalingDenom := udnScalingDenom; (* inc *)
stAxis.stScaling.lrScalingNum := lrScalingNum; (* deg *)
stAxis.stScaling.lrScaleFactor := udnScalingDenom / lrScalingNum;
stAxis.stPosition.lrOffsetPos := lrOriginShift;
stAxis.stLimitSwitches.lrSWPosLimitMin := lrSoftLimitMin;
stAxis.stLimitSwitches.lrSWPosLimitMax := lrSoftLimitMax;

A_AxisLink();
A_AxisGetStatus();
A_AxisController();
A_AxisMoveManual();
A_AxisMoveAuto();
A_AxisTerminalDiag();
A_AxisAlarm();


lrSpeedFactor := F_kAngleActuatorSpeedLin(
						bEnable := TRUE,
						lrActAngle := lrActPosition,
						lrAngleOffset := 56.6,  (* [deg] *)
						lrMultiplier := 0.755,
						lrOffset := 0.24
					);

Axis.stPlcToNc.stBaseDevice.stFastRefereneValue.nSpeed := LREAL_TO_INT(INT_TO_LREAL(Axis.stPlcToNc.stBaseDevice.stFastRefereneValue.nSpeed) * lrSpeedFactor);

*)

ACTION A_AxisAlarm:

(* Axis errors *)
tonAxisEnabled(
	IN := fbController.bEnable
		AND fbController.bRegulatorOn
		AND NOT fbController.bStatusDelay,
	PT := fbController.tStatusDelay + t#2s
);

bErrorCtrlEnabled := tonAxisEnabled.Q;
END_ACTION

ACTION A_AxisController:

(* Axis controller *)
fbController(
    bEnable := TRUE,
	etMachineMode := etMachineMode,
	etMachineState := etMachineState,
	bNoEStop := bNoEStop,
	bRegulatorOn := bNoEStop
				      AND bPowerSupplyOn
				      AND bSafetyOk
				      AND SEL(bNotMoving, NOT bCtrlInterrupt, TRUE)
				      AND NOT fbMoveManual.bControllerOff
				      AND NOT fbMoveAuto.bControllerOff,
	bReset := bConfirmAlarm,
	bTerminalOK := fbTerminalDiagnosis.bTerminalOK,
	bExeReset := bExeReset,
	bExeSetPos := FALSE,
	lrSetPosition := lrTargetPosition,
	bExeGearIn := bExeGearIn,
	bExeGearOut := bExeGearOut,
	dnRatioNumerator := dnRatioNumerator,
	udnRatioDenominator := udnRatioDenominator,
	lrOverride := SEL(bExtOverrideEn,
					lrOverride,
					lrOverride*lrExtOverride/100.0),
	bWithAbsoluteEncoder := bWithAbsoluteEncoder,
	bPosLagMonitoringEn := bPosLagMonitoringEn,
	lrPositionBias := 0.0,
	lrSoftLimitMax := lrSoftLimitMax,
	lrSoftLimitMin := lrSoftLimitMin,
	bSignalHWLimitMax:= bHWSignalLimitMax,
	bSignalHWLimitMin := bHWSignalLimitMin,
	lrAcceleration := lrAcceleration,
	lrDeceleration := lrDeceleration,
	lrJerk := lrJerk,
	pDrive := ADR(Drive),
	Axis := Axis,
	MasterAxis := MasterAxis,
	bStatusDelay => bCtrlEnabled,
	lrActPos => lrActPosition,
	lrActAbsPos => lrActAbsPosition,
	lrActVelo => lrActVelocity,
	bNotMoving => bNotMoving,
	bStandStill => bStandStill,
	bReferenced => bReferenced,
	bCoupled => bCoupled,
	lrVeloLimitMax => lrVeloMax,
	bHardLimitMaxExceeded => bHardLimitMaxExceeded,
	bHardLimitMinExceeded => bHardLimitMinExceeded,
	bSoftLimitMaxExceeded => bSoftLimitMaxExceeded,
	bSoftLimitMinExceeded => bSoftLimitMinExceeded
);

bSafetyDriveEnable := fbMoveManual.bSafetyCtrlEnable 
				 	  OR fbMoveAuto.bSafetyCtrlEnable;



(* from Tc2)

(* Axis controller *)
fbController(
    	bEnable := TRUE,
	etMachineMode := etMachineMode,
	etMachineState := etMachineState,
	bRegulatorOn := bNoEStop
				      AND bPowerSupplyOn
				      AND bSafetyOK
                 		      	      AND NOT bCtrlInterrupt
				      AND NOT fbMoveManual.bControllerOff
				      AND NOT fbMoveAuto.bControllerOff,
	bReset := bConfirmAlarm,
	bTerminalOK := fbTerminalDiagnosis.bTerminalOK,
	bExeReset := bExeReset,
	dwRawMotorEncoder := udnIncEnc,
	lrOverride := SEL(bExtOverrideEn,
					lrOverride,
					lrOverride*lrExtOverride/100.0),
	lrEngineTorque := SEL(
						bEngineTorqueLimitEn,
						nTorqueLimitMax,
						(lrEngineTorque) / 1),
	bWithAbsoluteEncoder := bWithAbsoluteEncoder,
	bHWSignalLimitMax := bHWSignalLimitMax,
	bHWSignalLimitMin := bHWSignalLimitMin,
	lrSoftLimitMax := lrSoftLimitMax,
	lrSoftLimitMin := lrSoftLimitMin,
	stEncoderConfig := stEncoderConfig,
	pAxis := ADR(stAxis),
	Axis := Axis,
	bStatusDelay => bCtrlEnabled,
	lrActPos=> ,
	lrActVelo => lrActVelocity,
	bNotMoving => bNotMoving,
	bReferenced => bReferenced,
	bHardLimitMaxExceeded => bHardLimitMaxExceeded,
	bHardLimitMinExceeded => bHardLimitMinExceeded,
	bSoftLimitMaxExceeded => bSoftLimitMaxExceeded,
	bSoftLimitMinExceeded => bSoftLimitMinExceeded
);

lrActPosition := F_LRealRound(fbController.lrActPos,1);
*)
END_ACTION

ACTION A_AxisGetStatus:

(* Get axis status *)
Axis.ReadStatus();
END_ACTION

ACTION A_AxisLink:

(* Get terminal status *)
sAdsAddr := F_CreateAmsNetId(Drive.stTerminalState.stAdsAddr.netId);
unSlaveAddr := Drive.stTerminalState.stAdsAddr.port;
Axis.DriveAddress.NetID := F_CreateAmsNetId(Drive.stTerminalState.stAdsAddr.netId);
Axis.DriveAddress.SlaveAddress := Drive.stTerminalState.stAdsAddr.port;

(* Set drive parameter *)
Drive.stPlcToStoeber.snA541ModesOfOperation := snModesOfOperation;

(*Drive.PlcToStoeber.nA558TargetTorque := SEL(bEngineTorqueLimitEn,
				    nTorqueLimitMax,
				    LREAL_TO_INT(lrEngineTorque / 1.0))*)
END_ACTION

ACTION A_AxisMoveAuto:

(* Move axis auto *)
rtMachineStandstill(CLK := bMachineStandstill);

lrVeloLimitMin := SEL(bVelocityLimitEn, -1 * lrVeloMax, lrVelocityMin);
lrVeloLimitMax := SEL(bVelocityLimitEn, lrVeloMax, lrVelocityMax);


fbMoveAuto(
	bEnable := bNoEStop
			   AND bPowerSupplyOn
			   AND bSafetyOK,
	bOccupied := bOccupied,
	bSafetyCtrlEnabled := bSafetyDriveEnabled,
	bCtrlEnabled := bCtrlEnabled
				      AND bMoveRelease,
	etMachineMode := etMachineMode,
	etMachineState := etMachineState,
	bReset := bConfirmAlarm,
	bCtrlEnable := bCtrlEnabled,
	bExeHome := bExeHome,
	bExeMoveAbs := bExeMoveAbs,
	bExeMoveVelo := bExeMoveVelo,
	bExeStop := bExeStop
			    OR rtMachineStandstill.Q,
	lrPosition := lrTargetPosition,
	lrVelocity := LIMIT(lrVeloLimitMin, lrAutoVelocity, lrVeloLimitMax),
	lrAcceleration := lrAcceleration,
	lrDeceleration := lrDeceleration,
	lrJerk := lrJerk,
	tControllerOff := tControllerOff,
	pDrive := ADR(Drive),
	bHomeCompleted := bHomeCompleted,
	Axis := Axis,
	MasterAxis := MasterAxis
 );
(* From Tc3) 

fbMoveAuto(
	bEnable := bNoEStop
               		    AND bPowerSupplyOn
               		    AND bSafetyOK,
	bCtrlEnabled := bCtrlEnabled
                    		   AND bMoveRelease,
	etMachineMode := etMachineMode,
	etMachineState := etMachineState,
	bReset := bConfirmAlarm,
	bExeHome := bExeHome,
	bExeMoveAbs := bExeMoveAbs,
	bExeMoveVelo := bExeMoveVelo,
	bExeStop := bExeStop
			      OR rtMachineStandstill.Q,
	lrPosition := lrTargetPosition,
	lrVelocity := LIMIT(lrVeloLimitMin, lrAutoVelocity, lrVeloLimitMax),
	lrAcceleration := lrAcceleration,
	lrDeceleration := lrDeceleration,
	lrJerk := lrJerk,
	tControllerOff := tControllerOff,
	stControllerConfig := stControllerConfig,
	pAxis := ADR(stAxis),
	bHomeCompleted := bHomeCompleted,
	Axis := Axis
 );
 
 *)
END_ACTION

ACTION A_AxisMoveManual:

(* Move axis manual *)
fbMoveManual(
	bEnable := bNoEStop
               		    AND bPowerSupplyOn
               		    AND bSafetyOK,
	bCtrlEnabled := bCtrlEnabled
               			    AND bMoveRelease,
	etMachineMode := etMachineMode,
	etMachineState := etMachineState,
	bReset := bConfirmAlarm,
	bMovePlus := bTipPlus,
	bMoveMinus := bTipMinus,
	bLimitMax := bHardLimitMaxExceeded
			       OR bSoftLimitMaxExceeded,
	bLimitMin := bHardLimitMinExceeded
			      OR bSoftLimitMinExceeded,
	bPlusRelease := bPlusRelease,
	bMinusRelease := bMinusRelease,
	lrVelocity := SEL(NOT bReferenced, lrManualVelocity, lrVelocityNoRef),
	tControllerOff := tControllerOff,
	bHomeCompleted := bHomeCompleted,
	Axis := Axis,
	MasterAxis 				:= GVL_Gr00Interface.iAxisDummy,
);

bSafetyLock := fbMoveManual.bMovePlus
                		OR fbMoveManual.bMoveMinus;
END_ACTION

ACTION A_AxisTerminalDiag:

(*Axis terminal diagnosis *)
fbTerminalDiagnosis(
	stTerminalState := Drive.stTerminalState,
	sTerminalStatus => sTerminalStatus
);

bErrorTerminal := NOT fbTerminalDiagnosis.bTerminalOK;
END_ACTION

END_FUNCTION_BLOCK

// ---- POUs/Tc2 Objects/MachineEquipment/F_kAngleActuatorSpeedLin.TcPOU
FUNCTION F_kAngleActuatorSpeedLin : LREAL
(*

The function used to linearization speed of angle actuator dependent of angle, sin()-function aligned 
Output factor: 0..1 (1=no speed reduction)

Constructor: 		Eduard Schüle
Company:		E. Riexinger GmbH
Date:			19.11.2015
Version:			1.00

Date:			Revision:		Who:				Comment
dd.mm.yyyy		x.xx			Initials			comment

*)
VAR_INPUT
	(* Input variables / Eingang Variablen *)
	bEnable							:BOOL;						(* Function block enable *)
	lrActAngle						:LREAL;						(* actual angle *)
	lrAngleOffset						:LREAL;						(* parameter sin-function angle offset *)
	lrMultiplier						:LREAL;						(* parameter sin-function multiplier *)
	lrOffset							:LREAL;						(* parameter sin-function offset *)
END_VAR
VAR
END_VAR

IF NOT bEnable
THEN
	F_kAngleActuatorSpeedLin := 1.0;
	RETURN;
END_IF

lrActAngle := LIMIT(-50, lrActAngle, 50);

F_kAngleActuatorSpeedLin := MIN(SIN( (lrActAngle + lrAngleOffset)/180*PI) * lrMultiplier + lrOffset, 1.0);

END_FUNCTION

// ---- POUs/Machine/Group_0100 - Production/Gr01Control/Gr01Alarm/FB_Gr01Alarm.TcPOU
FUNCTION_BLOCK FB_Gr01Alarm
(*

The function block used to control general alarms of machine.

Constructor: 		Patryk Panylo
Company:		E. Riexinger GmbH
Date:			28.04.2015
Version:			1.00

Date:			Revision:		Who:				Comment
dd.mm.yyyy		x.xx			Initials			comment

*)
VAR_INPUT
	(* Input variables / Eingang Variablen *)
	etMachineMode				:ET_MachineMode;			(* Machine mode *)
	etMachineState				:ET_MachineState;			(* Machine state *)
	bNoEStop					:BOOL;						(* Emergency stop *)
	bConfirmAlarm				:BOOL;						(* Confirm alarm *)
	dtDateTime 					:DATE_AND_TIME;			(* Actual date and time *)
	nFatalErrorMaxIdx				:INT;						(* Maximal index of  using alarms *)
	nErrorMaxIdx					:INT;						(* Maximal index of  using alarms *)
	nWarningMaxIdx				:INT;						(* Maximal index of  using alarms *)
	nMessageMaxIdx				:INT;						(* Maximal index of  using alarms *)
	nHintMaxIdx					:INT;						(* Maximal index of  using alarms *)
	stAlarmIn						:ST_AlarmIn;					(* Alarm input *)
END_VAR
VAR_OUTPUT
	(* Output variables / Ausgang Variablen *)
	stAlarmOut					:ST_AlarmOut;				(* Alarm input *)
END_VAR
VAR_IN_OUT
	(* Input Output variables / Ausgang Variablen *)
	bMoveInterrupted				:BOOL;						(* Move interrupted *)
	bHomeCompleted				:BOOL;						(* Home completed *)
END_VAR
VAR
	(* Enummerations *)

	(* Variables *)

	(* References *)

	(* Interfaces *)

	(* Instances *)
	fbAlarm						:FB_Alarm;
END_VAR


(* Collection of alarms *)
fbAlarm(
	bEnable := TRUE,
	bNoEStop := bNoEStop,
	bReset := bConfirmAlarm,
	dtDateTime := dtDateTime,
	nFatalErrorMaxIdx := nFatalErrorMaxIdx,
	nErrorMaxIdx := nErrorMaxIdx,
	nWarningMaxIdx := nWarningMaxIdx,
	nMessageMaxIdx := nMessageMaxIdx,
	nHintMaxIdx := nHintMaxIdx,
    	stAlarmIn := stAlarmIn,
    	stAlarmOut => stAlarmOut
);

IF stAlarmOut.bFatalError
    OR stAlarmOut.bError
THEN
	(*bMoveInterrupted := FALSE;*)
	bHomeCompleted := FALSE;
END_IF;

END_FUNCTION_BLOCK

// ---- POUs/Machine/Group_0100 - Production/Gr01Control/Gr01Safety/FB_Gr01Safety.TcPOU
FUNCTION_BLOCK FB_Gr01Safety
(*

The function block used to control genaeral safety of the machine.

Constructor: 		Patryk Panylo
Company:		E. Riexinger GmbH
Date:			28.04.2015
Version:			1.00

Date:			Revision:		Who:				Comment
dd.mm.yyyy		x.xx			Initials			comment

*)
VAR_INPUT
	(* Input variables / Eingang Variablen *)
	etMachineMode				:ET_MachineMode;			(* Machine mode *)
	etMachineState				:ET_MachineState;			(* Machine state *)
	bLightCurtain					:BOOL;						(* Light curtain ok / Freigabe Lichtschranke i.o *)
	bConfirmLightCurtain			:BOOL;						(* Confirm light Curtain input signal *)
	tLightCurtainDelay				:TIME := t#1s;					(* After time light Curtain safe *)
END_VAR
VAR_OUTPUT
	(* Output variables / Ausgang Variablen *)
	bLightCurtainOK				:BOOL;						(* Light curtain ok / Freigabe Lichtschranke i.o *)
	bConfirmedLightCurtain			:BOOL;						(* Confirmed light Curtain signal *)
	bNotInCrashArea				:BOOL;						(* Axis not in crash area with *)
	bPipeNotInCrashArea			:BOOL;						(* Axis not in crash with pipe *)
END_VAR
VAR_IN_OUT
	(* Input Output variables / Ausgang Variablen *)

END_VAR
VAR
	(* Enummerations *)

	(* Variables *)

	(* References *)

	(* Interfaces *)

	(* Instances *)
	fbLightCurtain					:FB_LightCurtain;

END_VAR


A_LightCurtain();
A_SafetyArea();

ACTION A_LightCurtain:

(* Light Curtain control *)
fbLightCurtain(
	bEnable := TRUE,
	bIn := bLightCurtain,
	bInConf := bConfirmLightCurtain,
	tTimeOut := tLightCurtainDelay,
	bOut => bLightCurtainOK,
	bOutConf => bConfirmedLightCurtain
);
END_ACTION

ACTION A_SafetyArea:

(* Safety area *)

bNotInCrashArea := FALSE;

IF FALSE
THEN
	bNotInCrashArea := TRUE;
END_IF;

IF bgGr01PipePresent
     (* AND NOT bgGr00ModeAutomatic*) 	(* 20260219 ES/KG *)
     AND MAX(0, stgGr01HMI.stPLCTOHMI.lrAxisSawBowActPos - lrgGr01DistSawbandPipe) > stgGr01HMI.stHMITOPLC.rPipeDiameter
     AND  Gr01Control.fbAxisSawBow.lrActVelocity < 0 		(* from Tc2) igGr01AxisSawBow.stNcToPlc.stBaseDevice.stCommandPositioning.dnActVelocity < 0 *)
THEN
	bPipeNotInCrashArea := FALSE;
ELSE
	bPipeNotInCrashArea := TRUE;
END_IF;
END_ACTION

END_FUNCTION_BLOCK

// ---- POUs/Machine/Group_0100 - Production/Gr01Control/Gr01Signals/FB_Gr01Signals.TcPOU
FUNCTION_BLOCK FB_Gr01Signals
(*

The function block used to control general signals of the machine.

Constructor: 		Patryk Panylo
Company:		E. Riexinger GmbH
Date:			28.04.2015
Version:			1.00

Date:			Revision:		Who:				Comment
dd.mm.yyyy		x.xx			Initials			comment

*)
VAR_INPUT
	(* Input variables / Eingang Variablen *)
	etMachineMode				:ET_MachineMode;			(* Machine mode *)
	etMachineState				:ET_MachineState;			(* Machine state *)
	bMachineRunning				:BOOL;						(* Machine running / Maschine lauft *)
	bExecutedProcess			:BOOL;						(* Process executed *)
	stBlinker						:ST_Blinker;
END_VAR
VAR_OUTPUT
	(* Output variables / Ausgang Variablen *)
	bBulbBtnStop					:BOOL;						(* Signal button bulb "stop" / Signallampe "Stop" *)
	bBulbBtnStart					:BOOL;						(* Signal button bulb "start" / Signallampe "Start" *)
END_VAR
VAR_IN_OUT
	(* Input Output variables / Ausgang Variablen *)

END_VAR
VAR
	(* Enummerations *)

	(* Variables *)

	(* References *)

	(* Interfaces *)

	(* Instances *)

END_VAR


A_SignalButton();

ACTION A_SignalButton:

(* Signal button bulb "stop" / Signallampe "Stop" *)
bBulbBtnStop := NOT bExecutedProcess;


(* Signal button bulb "start" / Signallampe "Start" *)
bBulbBtnStart := SEL(bExecutedProcess,
                           		     bMachineRunning AND stBlinker.Q1,
                           		     bMachineRunning);
END_ACTION

END_FUNCTION_BLOCK

// ---- POUs/Machine/Group_0100 - Production/Gr01Control/Gr01Utility/FB_Gr01Utility.TcPOU
FUNCTION_BLOCK FB_Gr01Utility
(*

The function block used to control general utility of the machine.

Constructor: 		Patryk Panylo
Company:		E. Riexinger GmbH
Date:			28.04.2015
Version:			1.00

Date:			Revision:		Who:				Comment
dd.mm.yyyy		x.xx			Initials			comment

*)
VAR_INPUT
	(* Input variables / Eingang Variablen *)
	etMachineMode				:ET_MachineMode;			(* Machine mode *)
	etMachineState				:ET_MachineState;			(* Machine state *)
	arbStartProcess				:ARRAY[1..3] OF BOOL;		(* Start process *)
	arbStopProcess				:ARRAY[1..3] OF BOOL;		(* Stop process *)
	arbSteppingProcess			:ARRAY[1..3] OF BOOL;		(* Stepping process *)
	bAutoCompleted				:BOOL;						(* Process completed *)
	bExeCounter					:BOOL;						(* Execute counter *)
	bLaserOnOff					:BOOL;						(* Laser on / off *)
	bStartTime					:BOOL;						(* Start measurement of cylce time *)
	bStopTime					:BOOL;						(* Stop measurement of cylce time *)
	bLifetimeOn					:BOOL;						(* Lifetime on *)
	bResetLifetimeAll				:BOOL; 						(* Reset all counters *)
	bResetLifetime				:BOOL;						(* Reset counter *)
	sLifetimeFilePath				:STRING;					(* File path for life time *)
	sLifetimeFileName			:STRING;					(* File name for life time *)
	bPipeIdentify					:BOOL;						(* Pipe identify *)
	rGlobalOverride				:REAL;						(* Global override *)
	tAdsTimeOut 					:TIME := t#2s;					(* Timout for ads commands *)
END_VAR
VAR_OUTPUT
	(* Output variables / Ausgang Variablen *)
	arbExeProcess				:ARRAY[1..3] OF BOOL;		(* Execute process *)
	rActOverride					:REAL;						(* Actual override *)
	lrLifetimeAll					:LREAL;						(* Lifetime all *)
	lrLifetimeAfterReset			:LREAL;						(* Lifetime after reset *)
	lrLifetimeAfterTrunOn			:LREAL;						(* Lifetime after turn on *)
	bLaserOn					:BOOL;						(* Laser on*)
	bPipePresent					:BOOL;						(* End present *)
END_VAR
VAR_IN_OUT
	(* Input Output variables / Ausgang Variablen *)
	bHomeCompleted				:BOOL;						(* Execute process *)
	rLocalOverride				:REAL;						(* Actual override *)
	udnCounterTotal				:UDINT;						(* Counter *)
END_VAR
VAR
	(* Enummerations *)

	(* Variables *)
	nIdxStartProcess				:INT;
	arudnCounterTotal				:ARRAY[0..1] OF UDINT;			(* Counter *)

	(* References *)

	(* Interfaces *)

	(* Instances *)
	arfbStartProcess				:ARRAY[1..3] OF FB_StartProcess;
	fbOverride					:FB_Override;
	fbOverrideSelection			:FB_OverrideSelection;
	fbLifetime					:FB_TimeHoursCounter;		(* Machine lifetime *)
	arfbCounter					:ARRAY[0..1] OF FB_Counter;
	arfbCylceTime				:ARRAY[0..1] OF FB_Timer;
	fbPipeIdentify					:FB_SignalHandlingEdge;
	fbLaserOnOff					:FB_SignalHandlingEdge;
END_VAR


A_StartProcess();
A_Override();
A_Counter();
A_CycleTime();
A_Laser();
A_PipeIdentify();

ACTION A_Counter:

(* Hours counter *)
fbLifetime(
	bEnable := TRUE,
	bDeleteAll := bResetLifetimeAll,
	sAmsNetId := sgAmsNetId,
	bCount := bLifetimeOn,
	bSave := FALSE,
	bReset := bResetLifetime,
	sFilePath := sLifetimeFilePath,
	sFileName := sLifetimeFileName,
	tSaveIntervall := t#8m,
	tTimeout := tAdsTimeOut,
	lrAllOverHours => lrLifetimeAll,
	lrAfterResetHours => lrLifetimeAfterReset,
	lrNoRetainHours => lrLifetimeAfterTrunOn,
 );

(* Counter *)
arfbCounter[0](
	bEnable := TRUE,
	bExecute := bExeCounter,
	bReset := arfbCounter[0].bOverflow,
	udnCounter := udnCounterTotal
);

arfbCounter[1](
	bEnable := TRUE,
	bExecute := bExeCounter,
	bReset := arfbCounter[1].bOverflow,
	udnCounter := arudnCounterTotal[1]
);
END_ACTION

ACTION A_CycleTime:

(* Cylce time *)
arfbCylceTime[0](
	bEnable := TRUE,
	bReset := FALSE,
	bStartStop := bStartTime
			        AND bgGr00ModeAutomatic,
	bStop := bStopTime
		        OR bgGr00MachineStandstill,
	tMaxTime := t#480m,
	stRefTime => ,
	stActTime => ,
	stRestTime =>
);

arfbCylceTime[1](
	bEnable := TRUE,
	bReset := FALSE,
	bStartStop := bStartTime
			        AND bgGr00ModeAutomatic,
	bStop := bStopTime
		        OR bgGr00MachineStandstill,
	tMaxTime := t#480m,
	stRefTime => ,
	stActTime => ,
	stRestTime =>
);
END_ACTION

ACTION A_Laser:

fbLaserOnOff(
	bEnable := TRUE,
	bIn := bLaserOnOff,
	tDelay := t#0ms,
);

IF fbLaserOnOff.bRisingEdge
THEN
	bLaserOn := NOT bLaserOn;
END_IF;
END_ACTION

ACTION A_Override:

(* Override control *)
fbOverrideSelection(
	bEnable := TRUE,
	rGlobalOverride := rGlobalOverride,
	rLocalOverride := rLocalOverride
);

fbOverride(
	bEnable := TRUE,
	bBypassAccDec := etMachineMode = ET_MachineMode_eManual,
	rSetOverride := fbOverrideSelection.rActOverride,
	rAcc := rgGr01AdsOverrideAcc,
	rDec := rgGr00AdsOverrideDec,
	rActOverride => rActOverride
);
END_ACTION

ACTION A_PipeIdentify:

fbPipeIdentify(
	bEnable := TRUE,
	bIn := bPipeIdentify,
	tDelay := t#100ms,
	bOut => bPipePresent
);
END_ACTION

ACTION A_StartProcess:

(* Start auto process *)

FOR nIdxStartProcess := 1 TO 3
DO
	arfbStartProcess[nIdxStartProcess](
		bEnable := etMachineMode = ET_MachineMode_eAutomatic
				    OR etMachineMode = ET_MachineMode_eCycle
				    OR etMachineMode = ET_MachineMode_eStepping,
		bStart := arbStartProcess[nIdxStartProcess],
		bStop := arbStopProcess[nIdxStartProcess],
		bDone := bAutoCompleted,
		bStepping := arbSteppingProcess[nIdxStartProcess],
		bHomeCompleted := bHomeCompleted,
		bStartProcess =>
	);

	arbExeProcess[nIdxStartProcess] := arfbStartProcess[nIdxStartProcess].bStartProcess;
END_FOR
END_ACTION

END_FUNCTION_BLOCK

// ---- POUs/Tc2 Objects/Automation/Process/FB_StartProcess.TcPOU
FUNCTION_BLOCK FB_StartProcess
(*

The function block used to control start process.

Constructor: 		Patryk Panylo
Company:		E. Riexinger GmbH
Date:			27.04.2015
Version:			1.00

Date:			Revision:		Who:				Comment
dd.mm.yyyy		x.xx			Initials			comment

*)
VAR_INPUT
	(* Input variables / Eingang Variablen *)
	bEnable						:BOOL;						(* Enable FB signal *)
	bStart						:BOOL;						(* Signal start *)
	bStop						:BOOL;						(* Signal stop *)
	bDone						:BOOL;						(* Signal done *)
	bStepping					:BOOL;						(* Stepping active *)
END_VAR
VAR_OUTPUT
	(* Output variables / Ausgang Variablen *)
	bStartProcess				:BOOL;						(* Start process *)
END_VAR
VAR_IN_OUT
	(* Input Output variables / Ausgang Variablen *)
	bHomeCompleted				:BOOL;			(* Home completed *)
END_VAR
VAR
	(* Enummerations *)

	(* Variables *)

	(* References *)

	(* Interfaces *)

	(* Instances *)
	rtStart						:R_TRIG;
END_VAR

IF NOT bEnable
THEN
	rtStart(CLK := FALSE);
	bStartProcess := FALSE;
	RETURN;
END_IF;


(* Start process with handshake *)
rtStart(CLK:= bStart);

IF (bDone
      OR bStop
      OR NOT bHomeCompleted)
    AND bStartProcess
THEN
	bStartProcess := FALSE;

ELSIF rtStart.Q
             AND NOT bStartProcess
THEN
	IF bStepping
	THEN
		 bStartProcess := rtStart.Q;
	ELSE
		bStartProcess := TRUE;
	END_IF;
END_IF;

END_FUNCTION_BLOCK

// ---- POUs/Tc2 Objects/Automation/Axis/Override/FB_OverrideSelection.TcPOU
FUNCTION_BLOCK FB_OverrideSelection
(*

The function block used to select override of axis.

Constructor: 		Patryk Panylo
Company:		E. Riexinger GmbH
Date:			23.04.2015
Version:			1.00

Date:			Revision:		Who:				Comment
dd.mm.yyyy		x.xx			Initials			comment

*)
VAR_INPUT
	(* Input variables / Eingang Variablen *)
	bEnable						:BOOL;						(* Signal FB enable *)
	rGlobalOverride				:REAL;						(* Global override *)
	rAcc							:REAL;						(* Accerlation of Override [%/s] *)
	rDec						:REAL;						(* Decerlation of Override [%/s] *)
END_VAR
VAR_OUTPUT
	(* Output variables / Ausgang Variablen *)
	rActOverride					:REAL;						(* Actual override *)
	bActGlobalOverride			:BOOL;						(* Actual override is global *)
	bActLocalOverride			:BOOL;						(* Actual override is local *)
END_VAR
VAR_IN_OUT
	(* Input Output variables / Ausgang Variablen *)
	rLocalOverride				:REAL;						(* Actual override *)
END_VAR
VAR
	(* Enummerations *)

	(* Variables *)
	rCacheGlobalOverride			:REAL;						(* Caches global override *)
	rCacheLocalOverride			:REAL;						(* Caches local override *)

	bFirstTime					:BOOL;						(* First run *)

	(* References *)

	(* Interfaces *)

	(* Instances *)
	tonChkCycleTime				:TON;						(* Check cycle time *)
END_VAR
VAR CONSTANT

END_VAR


IF NOT bEnable
THEN
	bFirstTime := FALSE;                               		(* Firstrun *)
	rActOverride := 0.0;                               		(* Override to set *)
	bActGlobalOverride := FALSE;                       	(* Actual override is global *)
	bActLocalOverride := FALSE;                       	(* Actual override is local *)
	RETURN;
END_IF;

IF NOT bFirstTime
THEN
	rCacheGlobalOverride := rGlobalOverride;          	(* Cache values *)
	rCacheLocalOverride := rLocalOverride;            		(* Cache values *)
	bActGlobalOverride := TRUE;                        			(* Actual override is global *)
	bActLocalOverride := FALSE;                       			(* Actual override is local *)
	bFirstTime := TRUE;                                				(* Firstrun *)
END_IF;

A_SelectLocal();
A_SelectGlobal();

ACTION A_SelectGlobal:

IF rCacheGlobalOverride <> rGlobalOverride
    OR rLocalOverride >= rGlobalOverride
THEN
	rCacheGlobalOverride := rGlobalOverride;
	rActOverride := rGlobalOverride;
	bActGlobalOverride := TRUE;                       	 		(* Actual override is global *)
	bActLocalOverride := FALSE;                        			(* Actual override is local *)
	rLocalOverride := rGlobalOverride;                		(* Set local Override *)
	rCacheLocalOverride := rGlobalOverride;           		(* Set local Override *)
END_IF;
END_ACTION

ACTION A_SelectLocal:

IF rCacheLocalOverride <> rLocalOverride
    AND rLocalOverride < rGlobalOverride
THEN
	rCacheLocalOverride := rLocalOverride;
	rActOverride := rLocalOverride;
	bActGlobalOverride := FALSE;                       			(* Actual override is global *)
	bActLocalOverride := TRUE;                        			(* Actual override is local *)
END_IF;
END_ACTION

END_FUNCTION_BLOCK

// ---- POUs/Tc2 Objects/Signals/Handling/FB_SignalHandlingEdge.TcPOU
FUNCTION_BLOCK FB_SignalHandlingEdge
VAR_INPUT
	(* Input variables / Eingang Variablen *)
	bEnable					:BOOL;						(* Enable FB signal *)
	bIn						:BOOL;						(* Input signal *)
	tDelay					:TIME := t#0s;					(* Delay *)
END_VAR
VAR_OUTPUT
	(* Output variables / Ausgang Variablen *)
	bOut					:BOOL;						(* Delayed signal *)
	bRisingEdge				:BOOL;						(* Rising edge *)
	bFallingEdge				:BOOL;						(* Falling edge *)
	bRisingEdgeDelay		:BOOL;						(* Rising edge delay *)
END_VAR
VAR
	(* Enummerations *)

	(* Variables *)


	(* References *)

	(* Interfaces *)

	(* Instances *)
	rtREdge					:R_TRIG;						(* Timer to delay *)
	rtREdgeDelay			:R_TRIG;						(* Timer to delay *)
	ftFEdge					:F_TRIG;						(* Timer to delay *)
	fbSignalHandlingDelay		:FB_SignalHandlingDelay;
END_VAR

IF NOT bEnable
THEN
	fbSignalHandlingDelay(
		bEnable := FALSE,
		bIn := bIn,
		bOut => bOut
	);

	rtREdge(CLK := FALSE);		(* Check rising edge *)
	ftFEdge(CLK := FALSE);		(* Check rising edge *)
	bRisingEdge := FALSE;
	bFallingEdge := FALSE;

	rtREdgeDelay(CLK := FALSE);		(* Check rising edge *)
	bRisingEdgeDelay := FALSE;
    RETURN;
END_IF;

fbSignalHandlingDelay(
	bEnable := TRUE,
	bIn := bIn,
	tDelay := tDelay,
	bOut => bOut
);

rtREdge(CLK := bIn);            			 (* Check rising edge *)
bRisingEdge := rtREdge.Q;

rtREdgeDelay(CLK := bOut);            			 (* Check rising edge *)
bRisingEdgeDelay := rtREdgeDelay.Q;

ftFEdge(CLK := bIn);            			 (* Check rising edge *)
bFallingEdge := ftFEdge.Q;

END_FUNCTION_BLOCK

// ---- POUs/Machine/Group_0100 - Production/Gr01MachineMode/Gr01Auto/Gr01Auto.TcPOU
PROGRAM Gr01Auto
VAR_INPUT
	(* Input variables / Eingang Variablen *)
	bEnable					:BOOL;						(* Enable Gr01Auto *)
	bExecute				:BOOL;						(* Auto execute *)

	(* Instances *)
	fbInit						:FB_Gr01AutoInit;
	fbProcedure				:FB_Gr01AutoProcedure;

END_VAR
VAR
	(* Enummerations *)

	(* Variables *)
	nIdx			:INT;

	(* References *)

	(* Interfaces *)

	(* Instances *)
	rtExecute					:R_TRIG;
	fbAlarm					:FB_Gr01AutoAlarm;
END_VAR
VAR CONSTANT
	nFatalErrorMaxIdx				:INT := 0;						(* Maximal index of  using alarms *)
	nErrorMaxIdx					:INT := 1;						(* Maximal index of  using alarms *)
	nWarningMaxIdx				:INT := 0;						(* Maximal index of  using alarms *)
	nMessageMaxIdx				:INT := 0;						(* Maximal index of  using alarms *)
	nHintMaxIdx					:INT := 0;						(* Maximal index of  using alarms *)

	dnFatalErrorBaseIdentNo		:DINT := 12000;				(* Fatal error identification number *)
	dnErrorBaseIdentNo			:DINT := 12100;				(* Error identification number *)
	dnWarningBaseIdentNo		:DINT := 12200;				(* Warning identification number *)
	dnMessageBaseIdentNo		:DINT := 12300;				(* Message identification number *)
	dnHintBaseIdentNo			:DINT := 12400;				(* Hint identification number *)
END_VAR

IF NOT bEnable
THEN
    RETURN;
END_IF;

(* Check auto execute *)
bExecute := bgGr00ModeAutomatic
		     AND NOT fbInit.bFirstTime;

rtExecute(CLK := bExecute);

IF rtExecute.Q
THEN
	A_Init();
END_IF;

A_Procedure();
A_Functions();
A_Alarm();

ACTION A_Alarm:

(* Collect and execute input alarms *)
fbAlarm.stAlarmIn.arbError[0].bActive := fbProcedure.bErrorCollisionDetected;
fbAlarm.stAlarmIn.arbError[0].dnCode := dnErrorBaseIdentNo + 0;

fbAlarm(
	etMachineMode := etgGr00MachineMode,
	etMachineState := etgGr00MachineState,
	bNoEStop := bgGr00NoEmergencyStop,
	bConfirmAlarm := bgGr00ConfirmAlarm,
	dtDateTime := stgGr00DateTime.dtDateTime,
	nFatalErrorMaxIdx := nFatalErrorMaxIdx,
	nErrorMaxIdx := nErrorMaxIdx,
	nWarningMaxIdx := nWarningMaxIdx,
	nMessageMaxIdx := nMessageMaxIdx,
	nHintMaxIdx := nHintMaxIdx,
	bMoveInterrupted := bgGr01MoveInterrupted,
	bHomeCompleted := bgGr01HomeCompleted,
	stAlarmOut => stgGr01Alarm.stAuto
);
END_ACTION

ACTION A_Functions:

;
END_ACTION

ACTION A_Init:

(* Initializing variables *)
fbInit();
END_ACTION

ACTION A_Procedure:

(* Execute auto procedure *)
fbProcedure(
	bEnable := fbInit.bFirstTime,
	bExecute := arbgGr01StartProcess[1]
			     OR arbgGr01StartProcess[2]
			     OR arbgGr01StartProcess[3],
	bInterrupt := FALSE(*NOT bgGr01StartProcess*),
	bReleaseNextStep := arbgGr01StartProcess[1]
					       OR arbgGr01StartProcess[2]
					       OR arbgGr01StartProcess[3],
	bDone => bgGr01AutoCompleted,
	bInterrupted => bgGr01MoveInterrupted
);
END_ACTION

END_PROGRAM

// ---- POUs/Tc2 Objects/Automation/Axis/F_ChkAllAxisEnabled.TcPOU
FUNCTION F_ChkAllAxisEnabled : BOOL
(*

The function used to detect if all axis controller enabled.

Constructor: 		Patryk Panylo
Company:		E. Riexinger GmbH
Date:			23.04.2015
Version:			1.00

Date:			Revision:		Who:				Comment
dd.mm.yyyy		x.xx			Initials			comment

*)
VAR_INPUT
	(* Input variables / Eingang Variablen *)
	bEnable						:BOOL;						(* Signal FB enable *)
	bEnabledAxis1				:BOOL;						(* Controller enabled *)
	bEnabledAxis2				:BOOL;						(* Controller enabled *)
	bEnabledAxis3				:BOOL;						(* Controller enabled *)
	bEnabledAxis4				:BOOL;						(* Controller enabled *)
	bEnabledAxis5				:BOOL;						(* Controller enabled *)
	bEnabledAxis6				:BOOL;						(* Controller enabled *)
	bEnabledAxis7				:BOOL;						(* Controller enabled *)
	bEnabledAxis8				:BOOL;						(* Controller enabled *)
	bEnabledAxis9				:BOOL;						(* Controller enabled *)
	bEnabledAxis10				:BOOL;						(* Controller enabled *)
END_VAR
VAR
	(* Enummerations *)

	(* Variables *)

	(* References *)

	(* Interfaces *)

	(* Instances *)

END_VAR


IF NOT bEnable							(* Signal FB enable *)
THEN
	F_ChkAllAxisEnabled := FALSE;

	RETURN;
END_IF

F_ChkAllAxisEnabled := bEnabledAxis1
					  AND bEnabledAxis2
					  AND bEnabledAxis3
					  AND bEnabledAxis4
					  AND bEnabledAxis5
					  AND bEnabledAxis6
					  AND bEnabledAxis7
					  AND bEnabledAxis8
					  AND bEnabledAxis9
					  AND bEnabledAxis10;

END_FUNCTION

// ---- POUs/Tc2 Objects/Automation/Axis/F_ChkAllAxisStandStill.TcPOU
FUNCTION F_ChkAllAxisStandStill : BOOL
(*

The function used to detect if all axis stand still.

Constructor: 		Patryk Panylo
Company:		E. Riexinger GmbH
Date:			23.04.2015
Version:			1.00

Date:			Revision:		Who:				Comment
dd.mm.yyyy		x.xx			Initials			comment

*)
VAR_INPUT
	(* Input variables / Eingang Variablen *)
	bEnable						:BOOL;					(* Signal FB enable *)
	bAxis1StandStill				:BOOL;					(* Axis stand still *)
	bAxis2StandStill				:BOOL;					(* Axis stand still *)
	bAxis3StandStill				:BOOL;					(* Axis stand still *)
	bAxis4StandStill				:BOOL;					(* Axis stand still *)
	bAxis5StandStill				:BOOL;					(* Axis stand still *)
	bAxis6StandStill				:BOOL;					(* Axis stand still *)
	bAxis7StandStill				:BOOL;					(* Axis stand still *)
	bAxis8StandStill				:BOOL;					(* Axis stand still *)
	bAxis9StandStill				:BOOL;					(* Axis stand still *)
	bAxis10StandStill				:BOOL;					(* Axis stand still *)
END_VAR
VAR
	(* Enummerations *)

	(* Variables *)

	(* References *)

	(* Interfaces *)

	(* Instances *)

END_VAR


IF NOT bEnable							(* Signal FB enable *)
THEN
	F_ChkAllAxisStandStill := FALSE;

	RETURN;
END_IF

F_ChkAllAxisStandStill := bAxis1StandStill
					   AND bAxis2StandStill
					   AND bAxis3StandStill
					   AND bAxis4StandStill
					   AND bAxis5StandStill
					   AND bAxis6StandStill
					   AND bAxis7StandStill
					   AND bAxis8StandStill
					   AND bAxis9StandStill
					   AND bAxis10StandStill;

END_FUNCTION

// ---- POUs/Tc2 Objects/Automation/Axis/F_ChkAllAxisNotMoving.TcPOU
FUNCTION F_ChkAllAxisNotMoving : BOOL
(*

The function used to detect if all axis not moving.

Constructor: 		Patryk Panylo
Company:		E. Riexinger GmbH
Date:			23.04.2015
Version:			1.00

Date:			Revision:		Who:				Comment
dd.mm.yyyy		x.xx			Initials			comment

*)
VAR_INPUT
	(* Input variables / Eingang Variablen *)
	bEnable						:BOOL;						(* Signal FB enable *)
	bAxis1NotMoving				:BOOL;						(* Axis not moving *)
	bAxis2NotMoving				:BOOL;						(* Axis not moving *)
	bAxis3NotMoving				:BOOL;						(* Axis not moving *)
	bAxis4NotMoving				:BOOL;						(* Axis not moving *)
	bAxis5NotMoving				:BOOL;						(* Axis not moving *)
	bAxis6NotMoving				:BOOL;						(* Axis not moving *)
	bAxis7NotMoving				:BOOL;						(* Axis not moving *)
	bAxis8NotMoving				:BOOL;						(* Axis not moving *)
	bAxis9NotMoving				:BOOL;						(* Axis not moving *)
	bAxis10NotMoving			:BOOL;						(* Axis not moving *)
END_VAR
VAR
	(* Enummerations *)

	(* Variables *)

	(* References *)

	(* Interfaces *)

	(* Instances *)

END_VAR


IF NOT bEnable							(* Signal FB enable *)
THEN
	F_ChkAllAxisNotMoving := FALSE;

	RETURN;
END_IF

F_ChkAllAxisNotMoving := bAxis1NotMoving
					   AND bAxis2NotMoving
					   AND bAxis3NotMoving
					   AND bAxis4NotMoving
					   AND bAxis5NotMoving
					   AND bAxis6NotMoving
					   AND bAxis7NotMoving
					   AND bAxis8NotMoving
					   AND bAxis9NotMoving
					   AND bAxis10NotMoving;

END_FUNCTION

// ---- POUs/Tc2 Objects/Automation/Axis/F_ChkAllAxisReferenced.TcPOU
FUNCTION F_ChkAllAxisReferenced : BOOL
(*

The function used to detect if all axis referenced.

Constructor: 		Patryk Panylo
Company:		E. Riexinger GmbH
Date:			23.04.2015
Version:			1.00

Date:			Revision:		Who:				Comment
dd.mm.yyyy		x.xx			Initials			comment

*)
VAR_INPUT
	(* Input variables / Eingang Variablen *)
	bEnable						:BOOL;						(* Signal FB enable *)
	bReferencedAxis1				:BOOL;						(* Controller referenced *)
	bReferencedAxis2				:BOOL;						(* Controller referenced *)
	bReferencedAxis3				:BOOL;						(* Controller referenced *)
	bReferencedAxis4				:BOOL;						(* Controller referenced *)
	bReferencedAxis5				:BOOL;						(* Controller referenced *)
	bReferencedAxis6				:BOOL;						(* Controller referenced *)
	bReferencedAxis7				:BOOL;						(* Controller referenced *)
	bReferencedAxis8				:BOOL;						(* Controller referenced *)
	bReferencedAxis9				:BOOL;						(* Controller referenced *)
	bReferencedAxis10			:BOOL;						(* Controller referenced *)
END_VAR
VAR
	(* Enummerations *)

	(* Variables *)

	(* References *)

	(* Interfaces *)

	(* Instances *)

END_VAR


IF NOT bEnable                          (* Signal FB enable *)
THEN
	F_ChkAllAxisReferenced := FALSE;

	RETURN;
END_IF;

F_ChkAllAxisReferenced := bReferencedAxis1
						AND bReferencedAxis2
						AND bReferencedAxis3
						AND bReferencedAxis4
						AND bReferencedAxis5
						AND bReferencedAxis6
						AND bReferencedAxis7
						AND bReferencedAxis8
						AND bReferencedAxis9
						AND bReferencedAxis10;

END_FUNCTION

// ---- POUs/Machine/Group_0000 - General/Gr00MachineMode/Gr00HMI/Gr00HMI.TcPOU
PROGRAM Gr00HMI
VAR_INPUT
	(* Input variables / Eingang Variablen *)
	bEnable					:BOOL;						(* Enable Gr00HMI *)
END_VAR
VAR
	(* Enummerations *)

	(* Variables *)

	(* References *)

	(* Interfaces *)

	(* Instances *)

END_VAR

IF NOT bEnable
THEN
	RETURN;
END_IF;

A_GetHMIVar();
A_SetHMIVar();

ACTION A_GetHMIVar:

(* Collect hmi signals *)
;
END_ACTION

ACTION A_SetHMIVar:

(* Collect hmi signals *)
stgGr00HMI.stPLCTOHMI.etMachineMode := etgGr00MachineMode;
stgGr00HMI.stPLCTOHMI.etMachineState := etgGr00MachineState;
stgGr00HMI.stPLCTOHMI.bHomeCompleted := bgGr00HomeCompleted;
stgGr00HMI.stPLCTOHMI.wBtnStartStatus.0 := bgGr00MachineRunning;
stgGr00HMI.stPLCTOHMI.wBtnStopStatus.0 := bgGr00MachineStandstill;
stgGr00HMI.stPLCTOHMI.wBtnResetStatus.0 := Gr00Control.fbSignals.stAlarm.bFatalError
                                                 					OR Gr00Control.fbSignals.stAlarm.bError
                                                					OR Gr00Control.fbSignals.stAlarm.bWarning;
stgGr00HMI.stPLCTOHMI.wBtnForceRefStatus.0 := Gr00Control.fbUtility.bSignalReference;
stgGr00HMI.stPLCTOHMI.bMachineRunning := bgGr00MachineRunning;
stgGr00HMI.stPLCTOHMI.bModeAutomatic := bgGr00ModeAutomatic;
stgGr00HMI.stPLCTOHMI.bModeHome := bgGr00ModeHome;
stgGr00HMI.stPLCTOHMI.bModeManual := bgGr00ModeManual;
stgGr00HMI.stPLCTOHMI.wAlarmStatus.0 := Gr00Control.fbSignals.stAlarm.bFatalError;
stgGr00HMI.stPLCTOHMI.wAlarmStatus.1 := Gr00Control.fbSignals.stAlarm.bError;
stgGr00HMI.stPLCTOHMI.wAlarmStatus.2 := Gr00Control.fbSignals.stAlarm.bWarning;
stgGr00HMI.stPLCTOHMI.wAlarmStatus.3 := Gr00Control.fbSignals.stAlarm.bMessage;
stgGr00HMI.stPLCTOHMI.wAlarmStatus.4 := Gr00Control.fbSignals.stAlarm.bHint;
stgGr00HMI.stPLCTOHMI.wLampStatus.0 := boutGr00BulbGreen;
stgGr00HMI.stPLCTOHMI.wLampStatus.1 := boutGr00BulbYellow;
stgGr00HMI.stPLCTOHMI.wLampStatus.2 := boutGr00BulbRed;
END_ACTION

END_PROGRAM

// ---- POUs/Machine/Group_0100 - Production/Gr01Coordinator.TcPOU
PROGRAM Gr01Coordinator
VAR_INPUT
	(* Input variables / Eingang Variablen *)
	bEnable					:BOOL;						(* Enable Group01 *)
END_VAR
VAR
	(* Enummerations *)

	(* Variables *)

	(* References *)

	(* Interfaces *)

	(* Instances *)

END_VAR

IF NOT bEnable
THEN
	RETURN;
END_IF;

Gr01Persistent(bEnable := TRUE);			(* Call Program *)
Gr01Simulation(bEnable := TRUE);			(* Call Program *)
Gr01MachineMode(bEnable := TRUE);		(* Call Program *)
Gr01Control(bEnable := TRUE);				(* Call Program *)
Gr01HMI(bEnable := TRUE);				(* Call Program *)

END_PROGRAM

// ---- POUs/Machine/Group_0100 - Production/Gr01Persistent/Gr01Persistent.TcPOU
PROGRAM Gr01Persistent
VAR_INPUT
	(* Input variables / Eingang Variablen *)
	bEnable								:BOOL;						(* Enable Gr01Persistent *)
END_VAR
VAR PERSISTENT
	(* Enummerations *)

	(* Variables *)
	rOverride							:REAL;											(* Override 0 - 100 [%]  *)
	udnCounterTotal						:UDINT;											(* Total counter *)

	lrAxisSawBowTipDistance				:LREAL;											(* Tip distance axis saw bow [mm] *)
	lrAxisSawBowOriginShiftPos			:LREAL;											(* Origin shift position axis saw bow [mm] *)
	lrAxisSawBowHomePos				:LREAL;											(* Home position axis saw bow [mm] *)
	lrAxisSawBowSoftLimitMax				:LREAL;											(* Software limit maximum axis saw bow [mm] *)
	lrAxisSawBowSoftLimitMin				:LREAL;											(* Software limit minimum axis saw bow [mm] *)
	lrAxisSawBowNoRefVelo				:LREAL;											(* No reference velocity axis saw bow [%] *)
	lrAxisSawBowManualVelo				:LREAL;											(* Manual velocity axis saw bow [%] *)
	lrAxisSawBowHomeVelo				:LREAL;											(* Home velocity axis saw bow [%] *)
	lrAxisSawBowAutoVelo					:LREAL;											(* Auto velocity axis saw bow [%] *)

	lrAxisAngleTipDistance				:LREAL;											(* Tip distance axis angle [mm] *)
	lrAxisAngleOriginShiftPos				:LREAL;											(* Origin shift position axis angle [mm] *)
	lrAxisAngleHomePos					:LREAL;											(* Home position axis angle [mm] *)
	lrAxisAngleSoftLimitMax				:LREAL;											(* Software limit maximum axis angle [mm] *)
	lrAxisAngleSoftLimitMin					:LREAL;											(* Software limit minimum axis angle [mm] *)
	lrAxisAngleNoRefVelo					:LREAL;											(* No reference velocity axis angle [mm/s] *)
	lrAxisAngleManualVelo					:LREAL;											(* Manual velocity axis angle [mm/s] *)
	lrAxisAngleHomeVelo					:LREAL;											(* Home velocity axis angle [mm/s] *)
	lrAxisAngleAutoVelo					:LREAL;											(* Auto velocity axis angle [mm/s] *)

	rSawbandManualSpeed				:REAL;											(* Manual speed sawband [upm] *)
	rSawbandAutoSpeed					:REAL;											(* Auto speed sawband [upm] *)
	rSawingOverride						:REAL;											(* Sawing override 0 - 100 [%]  *)
	rPipeDiameter						:REAL;											(* Pipe diameter [mm] *)
	lrActSawingAngle						:LREAL;											(* Actual angle of sawing [mm] *)
	lrSafetyDistance						:LREAL;											(* Safety distance [mm] *)
	lrSafeDistSawBandToPipe				:LREAL;											(* Safety distance sawband to pipe[mm] *)
	lrSawBandThickness					:LREAL;											(* Sawband thickness [mm] *)

	(* References *)

	(* Interfaces *)

	(* Instances *)
END_VAR
VAR
	(* Enummerations *)

	(* Variables *)
	bFirstTime							:BOOL;

	(* References *)

	(* Interfaces *)

	(* Instances *)

END_VAR

IF NOT bEnable
THEN
	bFirstTime := FALSE;
	RETURN;
END_IF;

IF NOT bFirstTime
THEN
	A_SetPerVar();

	bFirstTime := TRUE;
END_IF;

A_GetPerVar();

ACTION A_GetPerVar:

bgGr01WritePersistent := rOverride <> stgGr01HMI.stHMITOPLC.rOverride
					OR udnCounterTotal <> stgGr01HMI.stPLCTOHMI.udnCounterTotal
					OR lrAxisSawBowTipDistance <> stgGr01HMI.stHMITOPLC.lrAxisSawBowTipDistance
					OR lrAxisSawBowOriginShiftPos <> stgGr01HMI.stHMITOPLC.lrAxisSawBowOriginShiftPos
					OR lrAxisSawBowHomePos <> stgGr01HMI.stHMITOPLC.lrAxisSawBowHomePos
					OR lrAxisSawBowSoftLimitMax <> stgGr01HMI.stHMITOPLC.lrAxisSawBowSoftLimitMax
					OR lrAxisSawBowSoftLimitMin <> stgGr01HMI.stHMITOPLC.lrAxisSawBowSoftLimitMin
					OR lrAxisSawBowNoRefVelo <> stgGr01HMI.stHMITOPLC.lrAxisSawBowNoRefVelo
					OR lrAxisSawBowManualVelo <> stgGr01HMI.stHMITOPLC.lrAxisSawBowManualVelo
					OR lrAxisSawBowHomeVelo <> stgGr01HMI.stHMITOPLC.lrAxisSawBowHomeVelo
					OR lrAxisSawBowAutoVelo <> stgGr01HMI.stHMITOPLC.lrAxisSawBowAutoVelo

					OR lrAxisAngleTipDistance <> stgGr01HMI.stHMITOPLC.lrAxisAngleTipDistance
					OR lrAxisAngleOriginShiftPos <> stgGr01HMI.stHMITOPLC.lrAxisAngleOriginShiftPos
					OR lrAxisAngleHomePos <> stgGr01HMI.stHMITOPLC.lrAxisAngleHomePos
					OR lrAxisAngleSoftLimitMax <> stgGr01HMI.stHMITOPLC.lrAxisAngleSoftLimitMax
					OR lrAxisAngleSoftLimitMin <> stgGr01HMI.stHMITOPLC.lrAxisAngleSoftLimitMin
					OR lrAxisAngleNoRefVelo <> stgGr01HMI.stHMITOPLC.lrAxisAngleNoRefVelo
					OR lrAxisAngleManualVelo <> stgGr01HMI.stHMITOPLC.lrAxisAngleManualVelo
					OR lrAxisAngleHomeVelo <> stgGr01HMI.stHMITOPLC.lrAxisAngleHomeVelo
					OR lrAxisAngleAutoVelo <> stgGr01HMI.stHMITOPLC.lrAxisAngleAutoVelo

					OR rSawbandManualSpeed <> stgGr01HMI.stHMITOPLC.rSawbandManualSpeed
					OR rSawbandAutoSpeed <> stgGr01HMI.stHMITOPLC.rSawbandAutoSpeed
					OR rSawingOverride <> stgGr01HMI.stHMITOPLC.rSawingOverride
					OR rPipeDiameter <> stgGr01HMI.stHMITOPLC.rPipeDiameter
					OR lrActSawingAngle <> stgGr01HMI.stHMITOPLC.lrActSawingAngle
					OR lrSafetyDistance <> stgGr01HMI.stHMITOPLC.lrSafetyDistance
					OR lrSafeDistSawBandToPipe <> stgGr01HMI.stHMITOPLC.lrSafeDistSawBandToPipe
					OR lrSawBandThickness <> stgGr01HMI.stHMITOPLC.lrSawBandThickness;

rOverride := stgGr01HMI.stHMITOPLC.rOverride;
udnCounterTotal := stgGr01HMI.stPLCTOHMI.udnCounterTotal;

lrAxisSawBowTipDistance := stgGr01HMI.stHMITOPLC.lrAxisSawBowTipDistance;
lrAxisSawBowOriginShiftPos := stgGr01HMI.stHMITOPLC.lrAxisSawBowOriginShiftPos;
lrAxisSawBowHomePos := stgGr01HMI.stHMITOPLC.lrAxisSawBowHomePos;
lrAxisSawBowSoftLimitMax := stgGr01HMI.stHMITOPLC.lrAxisSawBowSoftLimitMax;
lrAxisSawBowSoftLimitMin := stgGr01HMI.stHMITOPLC.lrAxisSawBowSoftLimitMin;
lrAxisSawBowNoRefVelo := stgGr01HMI.stHMITOPLC.lrAxisSawBowNoRefVelo;
lrAxisSawBowManualVelo := stgGr01HMI.stHMITOPLC.lrAxisSawBowManualVelo;
lrAxisSawBowHomeVelo := stgGr01HMI.stHMITOPLC.lrAxisSawBowHomeVelo;
lrAxisSawBowAutoVelo := stgGr01HMI.stHMITOPLC.lrAxisSawBowAutoVelo;;

lrAxisAngleTipDistance := stgGr01HMI.stHMITOPLC.lrAxisAngleTipDistance;
lrAxisAngleOriginShiftPos := stgGr01HMI.stHMITOPLC.lrAxisAngleOriginShiftPos;
lrAxisAngleHomePos := stgGr01HMI.stHMITOPLC.lrAxisAngleHomePos;
lrAxisAngleSoftLimitMax := stgGr01HMI.stHMITOPLC.lrAxisAngleSoftLimitMax;
lrAxisAngleSoftLimitMin := stgGr01HMI.stHMITOPLC.lrAxisAngleSoftLimitMin;
lrAxisAngleNoRefVelo := stgGr01HMI.stHMITOPLC.lrAxisAngleNoRefVelo;
lrAxisAngleManualVelo := stgGr01HMI.stHMITOPLC.lrAxisAngleManualVelo;
lrAxisAngleHomeVelo := stgGr01HMI.stHMITOPLC.lrAxisAngleHomeVelo;
lrAxisAngleAutoVelo := stgGr01HMI.stHMITOPLC.lrAxisAngleAutoVelo;;

rSawbandManualSpeed := stgGr01HMI.stHMITOPLC.rSawbandManualSpeed;
rSawbandAutoSpeed := stgGr01HMI.stHMITOPLC.rSawbandAutoSpeed;
rSawingOverride := stgGr01HMI.stHMITOPLC.rSawingOverride;
rPipeDiameter := stgGr01HMI.stHMITOPLC.rPipeDiameter;
lrActSawingAngle := stgGr01HMI.stHMITOPLC.lrActSawingAngle;
lrSafetyDistance := stgGr01HMI.stHMITOPLC.lrSafetyDistance;
lrSafeDistSawBandToPipe := stgGr01HMI.stHMITOPLC.lrSafeDistSawBandToPipe;
lrSawBandThickness := stgGr01HMI.stHMITOPLC.lrSawBandThickness;
END_ACTION

ACTION A_SetPerVar:

stgGr01HMI.stHMITOPLC.rOverride := rOverride;
stgGr01HMI.stPLCTOHMI.udnCounterTotal := udnCounterTotal;

stgGr01HMI.stHMITOPLC.lrAxisSawBowTipDistance := lrAxisSawBowTipDistance;
stgGr01HMI.stHMITOPLC.lrAxisSawBowOriginShiftPos := lrAxisSawBowOriginShiftPos;
stgGr01HMI.stHMITOPLC.lrAxisSawBowHomePos := lrAxisSawBowHomePos;
stgGr01HMI.stHMITOPLC.lrAxisSawBowSoftLimitMax := lrAxisSawBowSoftLimitMax;
stgGr01HMI.stHMITOPLC.lrAxisSawBowSoftLimitMin := lrAxisSawBowSoftLimitMin;
stgGr01HMI.stHMITOPLC.lrAxisSawBowNoRefVelo := lrAxisSawBowNoRefVelo;
stgGr01HMI.stHMITOPLC.lrAxisSawBowManualVelo := lrAxisSawBowManualVelo;
stgGr01HMI.stHMITOPLC.lrAxisSawBowHomeVelo := lrAxisSawBowHomeVelo;
stgGr01HMI.stHMITOPLC.lrAxisSawBowAutoVelo := lrAxisSawBowAutoVelo;

stgGr01HMI.stHMITOPLC.lrAxisAngleTipDistance := lrAxisAngleTipDistance;
stgGr01HMI.stHMITOPLC.lrAxisAngleOriginShiftPos := lrAxisAngleOriginShiftPos;
stgGr01HMI.stHMITOPLC.lrAxisAngleHomePos := lrAxisAngleHomePos;
stgGr01HMI.stHMITOPLC.lrAxisAngleSoftLimitMax := lrAxisAngleSoftLimitMax;
stgGr01HMI.stHMITOPLC.lrAxisAngleSoftLimitMin := lrAxisAngleSoftLimitMin;
stgGr01HMI.stHMITOPLC.lrAxisAngleNoRefVelo := lrAxisAngleNoRefVelo;
stgGr01HMI.stHMITOPLC.lrAxisAngleManualVelo := lrAxisAngleManualVelo;
stgGr01HMI.stHMITOPLC.lrAxisAngleHomeVelo := lrAxisAngleHomeVelo;
stgGr01HMI.stHMITOPLC.lrAxisAngleAutoVelo := lrAxisAngleAutoVelo;

stgGr01HMI.stHMITOPLC.rSawbandManualSpeed := rSawbandManualSpeed;
stgGr01HMI.stHMITOPLC.rSawbandAutoSpeed := rSawbandAutoSpeed;
stgGr01HMI.stHMITOPLC.rSawingOverride := rSawingOverride;
stgGr01HMI.stHMITOPLC.rPipeDiameter := rPipeDiameter;
stgGr01HMI.stHMITOPLC.lrActSawingAngle := lrActSawingAngle;
stgGr01HMI.stHMITOPLC.lrSafetyDistance := lrSafetyDistance;
stgGr01HMI.stHMITOPLC.lrSafeDistSawBandToPipe := lrSafeDistSawBandToPipe;
stgGr01HMI.stHMITOPLC.lrSawBandThickness := lrSawBandThickness;
END_ACTION

END_PROGRAM

// ---- POUs/Machine/Group_0100 - Production/Gr01Simulation/Gr01Simulation.TcPOU
PROGRAM Gr01Simulation
VAR_INPUT
	(* Input variables / Eingang Variablen *)
	bEnable								:BOOL;						(* Enable Gr05Persistent *)
END_VAR
VAR
	(* Enummerations *)

	(* Variables *)

	(* References *)

	(* Interfaces *)

	(* Instances *)
END_VAR

IF NOT bEnable
THEN

	RETURN;
END_IF;

A_ForceInput();

ACTION A_ForceInput:


GVL_Gr00IO.binGr00AirPressureOK := TRUE;
GVL_Gr00IO.binGr00LightCurtainOK := TRUE;
GVL_Gr00IO.arbinGr00PowerSupplyOn[2] := TRUE;
GVL_Gr00IO.arbinGr00PowerSupplyOn[3] := TRUE;
GVL_Gr00IO.arbinGr00PowerSupplyOn[4] := TRUE;
GVL_Gr00IO.arbinGr00PowerSupplyOn[5] := TRUE;
GVL_Gr00IO.arbinGr00DoorsClosed[1] := TRUE;
GVL_Gr00IO.arbinGr00DoorsClosed[2] := TRUE;
GVL_Gr00IO.arbinGr00DoorsClosed[3] := TRUE;
GVL_Gr00IO.arbinGr00DoorsClosed[4] := TRUE;
GVL_Gr00IO.arbinGr00DoorsClosed[5] := TRUE;
GVL_Gr00IO.binGr00AllDoorsClosed := GVL_Gr00IO.arbinGr00DoorsClosed[1]
								AND GVL_Gr00IO.arbinGr00DoorsClosed[2]
								AND GVL_Gr00IO.arbinGr00DoorsClosed[3]
								AND GVL_Gr00IO.arbinGr00DoorsClosed[4]
								AND GVL_Gr00IO.arbinGr00DoorsClosed[5];

GVL_Gr00IO.binGr00AllDoorsLocked := TRUE;
GVL_Gr00IO.binGr00TempOK := TRUE;


// only for simulation
// GVL_Gr00IO.binNoEmergencyStop := TRUE;
// GVL_Gr00IO.binMoveRelease := TRUE;
// GVL_Gr00IO.binMoveReleaseSB := TRUE;
END_ACTION

END_PROGRAM

// ---- POUs/Machine/Group_0100 - Production/Gr01MachineMode/Gr01MachineMode.TcPOU
PROGRAM Gr01MachineMode
VAR_INPUT
	(* Input variables / Eingang Variablen *)
	bEnable					:BOOL;						(* Enable Gr01MachineMode *)
END_VAR
VAR
	(* Enummerations *)

	(* Variables *)

	(* References *)

	(* Interfaces *)

	(* Instances *)

END_VAR

IF NOT bEnable
THEN
	RETURN;
END_IF;

Gr01Auto(bEnable := TRUE);			(* Call Program *)
Gr01Home(bEnable := TRUE);			(* Call Program *)
Gr01Manual(bEnable := TRUE);			(* Call Program *)

END_PROGRAM

// ---- POUs/Machine/Group_0100 - Production/Gr01MachineMode/Gr01Manual/Gr01Manual.TcPOU
PROGRAM Gr01Manual
VAR_INPUT
	(* Input variables / Eingang Variablen *)
	bEnable					:BOOL;						(* Enable Gr01Manual *)
	bExecute				:BOOL;						(* Manual execute *)

	(* Instances *)
	fbInit						:FB_Gr01ManualInit;
	fbProcedure				:FB_Gr01ManualProcedure;
END_VAR
VAR
	(* Enummerations *)

	(* Variables *)

	(* References *)

	(* Interfaces *)

	(* Instances *)
	rtExecute					:R_TRIG;

	fbAlarm					:FB_Gr01ManualAlarm;
END_VAR
VAR CONSTANT
	nFatalErrorMaxIdx				:INT := 0;						(* Maximal index of  using alarms *)
	nErrorMaxIdx					:INT := 0;						(* Maximal index of  using alarms *)
	nWarningMaxIdx				:INT := 0;						(* Maximal index of  using alarms *)
	nMessageMaxIdx				:INT := 0;						(* Maximal index of  using alarms *)
	nHintMaxIdx					:INT := 0;						(* Maximal index of  using alarms *)

	dnFatalErrorBaseIdentNo		:DINT := 14000;				(* Fatal error identification number *)
	dnErrorBaseIdentNo			:DINT := 14100;				(* Error identification number *)
	dnWarningBaseIdentNo		:DINT := 14200;				(* Warning identification number *)
	dnMessageBaseIdentNo		:DINT := 14300;				(* Message identification number *)
	dnHintBaseIdentNo			:DINT := 14400;				(* Hint identification number *)
END_VAR

IF NOT bEnable
THEN
	RETURN;
END_IF;

(* Check manual execute *)
bExecute := etgGr00MachineMode = ET_MachineMode_eManual;

rtExecute(CLK := bExecute);

IF rtExecute.Q
THEN
	fbInit.bFirstTime := FALSE;
	A_Init();
END_IF;

A_Procedure();
A_Alarm();

ACTION A_Alarm:

(* Collect and execute input alarms *)
fbAlarm.stAlarmIn.arbError[0].bActive := FALSE;
fbAlarm.stAlarmIn.arbError[0].dnCode := dnErrorBaseIdentNo + 0;

fbAlarm(
	etMachineMode := etgGr00MachineMode,
	etMachineState := etgGr00MachineState,
	bNoEStop := bgGr00NoEmergencyStop,
	bConfirmAlarm := bgGr00ConfirmAlarm,
	dtDateTime := stgGr00DateTime.dtDateTime,
	nFatalErrorMaxIdx := nFatalErrorMaxIdx,
	nErrorMaxIdx := nErrorMaxIdx,
	nWarningMaxIdx := nWarningMaxIdx,
	nMessageMaxIdx := nMessageMaxIdx,
	nHintMaxIdx := nHintMaxIdx,
	bHomeCompleted := bgGr01HomeCompleted,
	stAlarmOut => stgGr01Alarm.stManual
);
END_ACTION

ACTION A_Init:

(* Initializing variables *)
fbInit();
END_ACTION

ACTION A_Procedure:

(* Execute manual procedure *)
fbProcedure(
	bEnable := etgGr00MachineMode = ET_MachineMode_eManual,
	bExecute := rtExecute.Q,
	bReleaseNextStep := etgGr00MachineMode = ET_MachineMode_eManual
);

IF fbProcedure.bDone
THEN
	bgGr01ManualCompleted := TRUE;
END_IF
END_ACTION

END_PROGRAM

// ---- POUs/Machine/Group_0100 - Production/Gr01HMI/Gr01HMI.TcPOU
PROGRAM Gr01HMI
VAR_INPUT
	(* Input variables / Eingang Variablen *)
	bEnable					:BOOL;						(* Enable Gr01HMI *)
END_VAR
VAR
	(* Enummerations *)

	(* Variables *)
	nIdx						:INT;

	(* References *)

	(* Interfaces *)

	(* Instances *)

END_VAR

IF NOT bEnable
THEN
	RETURN;
END_IF;

A_GetHMIVar();
A_SetHMIVar();

ACTION A_GetHMIVar:

(* Collect hmi signals *)
;
END_ACTION

ACTION A_SetHMIVar:

(* Collect hmi signals *)
stgGr01HMI.stPLCTOHMI.bHomeCompleted := bgGr01HomeCompleted;
stgGr01HMI.stPLCTOHMI.wBtnStartStatus.0 := arbgGr01StartProcess[1]
									       OR arbgGr01StartProcess[2]
									       OR arbgGr01StartProcess[3];
stgGr01HMI.stPLCTOHMI.wBtnStopStatus.0 := NOT arbgGr01StartProcess[1]
									       AND NOT arbgGr01StartProcess[2]
									       AND NOT arbgGr01StartProcess[3];
stgGr01HMI.stPLCTOHMI.wBtnStepProcStatus := 0;
stgGr01HMI.stPLCTOHMI.wAxisSawBowStatus.0 := NOT binGr01AxisSawBowLimitMin;
stgGr01HMI.stPLCTOHMI.wAxisSawBowStatus.1 := NOT binGr01AxisSawBowLimitMax;
stgGr01HMI.stPLCTOHMI.wAxisAngleStatus.0 := NOT binGr01AxisAngleLimitMin;
stgGr01HMI.stPLCTOHMI.wAxisAngleStatus.1 := NOT binGr01AxisAngleLimitMax;;
stgGr01HMI.stPLCTOHMI.wSawbandStatus.0 := FALSE;
stgGr01HMI.stPLCTOHMI.wSawbandStatus.1 := FALSE;
stgGr01HMI.stPLCTOHMI.wSawbandAirStatus.0 := boutGr01SawbandAirOn;
stgGr01HMI.stPLCTOHMI.wSawbandAirStatus.1 := NOT boutGr01SawbandAirOn;
stgGr01HMI.stPLCTOHMI.wLaserStatus.0 := boutGr01LaserOn;
stgGr01HMI.stPLCTOHMI.wLaserStatus.1 := NOT boutGr01LaserOn;
END_ACTION

END_PROGRAM

// ---- POUs/Machine/Group_0500 - Transport/Gr05Coordinator.TcPOU
PROGRAM Gr05Coordinator
VAR_INPUT
	(* Input variables / Eingang Variablen *)
	bEnable					:BOOL;						(* Enable Group05 *)
END_VAR
VAR
	(* Enummerations *)

	(* Variables *)

	(* References *)

	(* Interfaces *)

	(* Instances *)

END_VAR

IF NOT bEnable
THEN
	RETURN;
END_IF;

Gr05Persistent(bEnable := TRUE);			(* Call Program *)
Gr05Simulation(bEnable := TRUE);			(* Call Program *)
Gr05MachineMode(bEnable := TRUE);		(* Call Program *)
Gr05Control(bEnable := TRUE);				(* Call Program *)
Gr05HMI(bEnable := TRUE);				(* Call Program *)

END_PROGRAM

// ---- POUs/Machine/Group_0500 - Transport/Gr05Persistent/Gr05Persistent.TcPOU
PROGRAM Gr05Persistent
VAR_INPUT
	(* Input variables / Eingang Variablen *)
	bEnable								:BOOL;						(* Enable Gr05Persistent *)
END_VAR
VAR PERSISTENT
	(* Enummerations *)

	(* Variables *)
	rOverride							:REAL;						(* Override 0 - 100 % *)
	udnCounterTotal						:UDINT;						(* Total counter *)

	bSlideActive							:BOOL;											(* Slide active *)
	bCylinderPosActive					:BOOL;											(* Position cylinder active *)
	arlrAxisClampTipDistance				:ARRAY[1..ungGr05ClampMaxNo] OF LREAL;			(* Tip distance axis clamp [mm] *)
	arlrAxisClampOriginShiftPos				:ARRAY[1..ungGr05ClampMaxNo] OF LREAL;			(* Origin shift position axis clamp [mm] *)
	arlrAxisClampHomePos				:ARRAY[1..ungGr05ClampMaxNo] OF LREAL;			(* Home position axis clamp [mm] *)
	arlrAxisClampSoftLimitMax				:ARRAY[1..ungGr05ClampMaxNo] OF LREAL;			(* Software limit maximum axis clamp [mm] *)
	arlrAxisClampSoftLimitMin				:ARRAY[1..ungGr05ClampMaxNo] OF LREAL;			(* Software limit minimum axis clamp [mm] *)
	arlrAxisClampNoRefVelo				:ARRAY[1..ungGr05ClampMaxNo] OF LREAL;			(* No reference velocity axis clamp [mm/s] *)
	arlrAxisClampManualVelo				:ARRAY[1..ungGr05ClampMaxNo] OF LREAL;			(* Manual velocity axis clamp [mm/s] *)
	arlrAxisClampHomeVelo				:ARRAY[1..ungGr05ClampMaxNo] OF LREAL;			(* Home velocity axis clamp [mm/s] *)
	arlrAxisClampAutoVelo					:ARRAY[1..ungGr05ClampMaxNo] OF LREAL;			(* Auto velocity axis clamp [mm/s] *)
	lrActSawingLength						:LREAL;

	(* References *)

	(* Interfaces *)

	(* Instances *)
END_VAR
VAR
	(* Enummerations *)

	(* Variables *)
	bFirstTime							:BOOL;

	(* References *)

	(* Interfaces *)

	(* Instances *)

END_VAR

IF NOT bEnable
THEN
	bFirstTime := FALSE;
	RETURN;
END_IF;

IF NOT bFirstTime
THEN
	A_SetPerVar();

	bFirstTime := TRUE;
END_IF;

A_GetPerVar();

ACTION A_GetPerVar:

bgGr05WritePersistent := rOverride <> stgGr05HMI.stHMITOPLC.rOverride
					OR udnCounterTotal <> stgGr05HMI.stPLCTOHMI.udnCounterTotal
					OR bSlideActive <> stgGr05HMI.stHMITOPLC.bSlideActive
					OR bCylinderPosActive <> stgGr05HMI.stHMITOPLC.bCylinderPosActive
					OR MEMCMP(ADR(arlrAxisClampTipDistance), ADR(stgGr05HMI.stHMITOPLC.arlrAxisClampTipDistance), SIZEOF(stgGr05HMI.stHMITOPLC.arlrAxisClampTipDistance)) <> 0
					OR MEMCMP(ADR(arlrAxisClampOriginShiftPos), ADR(stgGr05HMI.stHMITOPLC.arlrAxisClampOriginShiftPos), SIZEOF(stgGr05HMI.stHMITOPLC.arlrAxisClampOriginShiftPos)) <> 0
					OR MEMCMP(ADR(arlrAxisClampHomePos), ADR(stgGr05HMI.stHMITOPLC.arlrAxisClampHomePos), SIZEOF(stgGr05HMI.stHMITOPLC.arlrAxisClampHomePos)) <> 0
					OR MEMCMP(ADR(arlrAxisClampSoftLimitMax), ADR(stgGr05HMI.stHMITOPLC.arlrAxisClampSoftLimitMax), SIZEOF(stgGr05HMI.stHMITOPLC.arlrAxisClampSoftLimitMax)) <> 0
					OR MEMCMP(ADR(arlrAxisClampSoftLimitMin), ADR(stgGr05HMI.stHMITOPLC.arlrAxisClampSoftLimitMin), SIZEOF(stgGr05HMI.stHMITOPLC.arlrAxisClampSoftLimitMin)) <> 0
					OR MEMCMP(ADR(arlrAxisClampNoRefVelo), ADR(stgGr05HMI.stHMITOPLC.arlrAxisClampNoRefVelo), SIZEOF(stgGr05HMI.stHMITOPLC.arlrAxisClampNoRefVelo)) <> 0
					OR MEMCMP(ADR(arlrAxisClampManualVelo), ADR(stgGr05HMI.stHMITOPLC.arlrAxisClampManualVelo), SIZEOF(stgGr05HMI.stHMITOPLC.arlrAxisClampManualVelo)) <> 0
					OR MEMCMP(ADR(arlrAxisClampHomeVelo), ADR(stgGr05HMI.stHMITOPLC.arlrAxisClampHomeVelo), SIZEOF(stgGr05HMI.stHMITOPLC.arlrAxisClampHomeVelo)) <> 0
					OR MEMCMP(ADR(arlrAxisClampAutoVelo), ADR(stgGr05HMI.stHMITOPLC.arlrAxisClampAutoVelo), SIZEOF(stgGr05HMI.stHMITOPLC.arlrAxisClampAutoVelo)) <> 0
					OR lrActSawingLength <> stgGr05HMI.stHMITOPLC.lrActSawingLength;


rOverride := stgGr05HMI.stHMITOPLC.rOverride;
udnCounterTotal := stgGr05HMI.stPLCTOHMI.udnCounterTotal;

bSlideActive := stgGr05HMI.stHMITOPLC.bSlideActive;
bCylinderPosActive := stgGr05HMI.stHMITOPLC.bCylinderPosActive;

MEMCPY(ADR(arlrAxisClampTipDistance), ADR(stgGr05HMI.stHMITOPLC.arlrAxisClampTipDistance), SIZEOF(stgGr05HMI.stHMITOPLC.arlrAxisClampTipDistance));
MEMCPY(ADR(arlrAxisClampOriginShiftPos), ADR(stgGr05HMI.stHMITOPLC.arlrAxisClampOriginShiftPos), SIZEOF(stgGr05HMI.stHMITOPLC.arlrAxisClampOriginShiftPos));
MEMCPY(ADR(arlrAxisClampHomePos), ADR(stgGr05HMI.stHMITOPLC.arlrAxisClampHomePos), SIZEOF(stgGr05HMI.stHMITOPLC.arlrAxisClampHomePos));
MEMCPY(ADR(arlrAxisClampSoftLimitMax), ADR(stgGr05HMI.stHMITOPLC.arlrAxisClampSoftLimitMax), SIZEOF(stgGr05HMI.stHMITOPLC.arlrAxisClampSoftLimitMax));
MEMCPY(ADR(arlrAxisClampSoftLimitMin), ADR(stgGr05HMI.stHMITOPLC.arlrAxisClampSoftLimitMin), SIZEOF(stgGr05HMI.stHMITOPLC.arlrAxisClampSoftLimitMin));
MEMCPY(ADR(arlrAxisClampNoRefVelo), ADR(stgGr05HMI.stHMITOPLC.arlrAxisClampNoRefVelo), SIZEOF(stgGr05HMI.stHMITOPLC.arlrAxisClampNoRefVelo));
MEMCPY(ADR(arlrAxisClampManualVelo), ADR(stgGr05HMI.stHMITOPLC.arlrAxisClampManualVelo), SIZEOF(stgGr05HMI.stHMITOPLC.arlrAxisClampManualVelo));
MEMCPY(ADR(arlrAxisClampHomeVelo), ADR(stgGr05HMI.stHMITOPLC.arlrAxisClampHomeVelo), SIZEOF(stgGr05HMI.stHMITOPLC.arlrAxisClampHomeVelo));
MEMCPY(ADR(arlrAxisClampAutoVelo), ADR(stgGr05HMI.stHMITOPLC.arlrAxisClampAutoVelo), SIZEOF(stgGr05HMI.stHMITOPLC.arlrAxisClampAutoVelo));

lrActSawingLength := stgGr05HMI.stHMITOPLC.lrActSawingLength;
END_ACTION

ACTION A_SetPerVar:

stgGr05HMI.stHMITOPLC.rOverride := rOverride;
stgGr05HMI.stPLCTOHMI.udnCounterTotal := udnCounterTotal;

stgGr05HMI.stHMITOPLC.bSlideActive := bSlideActive;
stgGr05HMI.stHMITOPLC.bCylinderPosActive := bCylinderPosActive;

MEMCPY(ADR(stgGr05HMI.stHMITOPLC.arlrAxisClampTipDistance), ADR(arlrAxisClampTipDistance), SIZEOF(arlrAxisClampTipDistance));
MEMCPY(ADR(stgGr05HMI.stHMITOPLC.arlrAxisClampOriginShiftPos), ADR(arlrAxisClampOriginShiftPos), SIZEOF(arlrAxisClampOriginShiftPos));
MEMCPY(ADR(stgGr05HMI.stHMITOPLC.arlrAxisClampHomePos), ADR(arlrAxisClampHomePos), SIZEOF(arlrAxisClampHomePos));
MEMCPY(ADR(stgGr05HMI.stHMITOPLC.arlrAxisClampSoftLimitMax), ADR(arlrAxisClampSoftLimitMax), SIZEOF(arlrAxisClampSoftLimitMax));
MEMCPY(ADR(stgGr05HMI.stHMITOPLC.arlrAxisClampSoftLimitMin), ADR(arlrAxisClampSoftLimitMin), SIZEOF(arlrAxisClampSoftLimitMin));
MEMCPY(ADR(stgGr05HMI.stHMITOPLC.arlrAxisClampNoRefVelo), ADR(arlrAxisClampNoRefVelo), SIZEOF(arlrAxisClampNoRefVelo));
MEMCPY(ADR(stgGr05HMI.stHMITOPLC.arlrAxisClampManualVelo), ADR(arlrAxisClampManualVelo), SIZEOF(arlrAxisClampManualVelo));
MEMCPY(ADR(stgGr05HMI.stHMITOPLC.arlrAxisClampHomeVelo), ADR(arlrAxisClampHomeVelo), SIZEOF(arlrAxisClampHomeVelo));
MEMCPY(ADR(stgGr05HMI.stHMITOPLC.arlrAxisClampAutoVelo), ADR(arlrAxisClampAutoVelo), SIZEOF(arlrAxisClampAutoVelo));

stgGr05HMI.stHMITOPLC.lrActSawingLength := lrActSawingLength;
END_ACTION

END_PROGRAM

// ---- POUs/Machine/Group_0500 - Transport/Gr05Simulation/Gr05Simulation.TcPOU
PROGRAM Gr05Simulation
VAR_INPUT
	(* Input variables / Eingang Variablen *)
	bEnable								:BOOL;						(* Enable Gr05Persistent *)
END_VAR
VAR
	(* Enummerations *)

	(* Variables *)

	(* References *)

	(* Interfaces *)

	(* Instances *)

END_VAR

IF NOT bEnable
THEN

	RETURN;
END_IF;

A_ForceInput();

ACTION A_ForceInput:


GVL_Gr00IO.binGr00AirPressureOK := TRUE;
GVL_Gr00IO.binGr00LightCurtainOK := TRUE;
GVL_Gr00IO.arbinGr00PowerSupplyOn[2] := TRUE;
GVL_Gr00IO.arbinGr00PowerSupplyOn[3] := TRUE;
GVL_Gr00IO.arbinGr00PowerSupplyOn[4] := TRUE;
GVL_Gr00IO.arbinGr00PowerSupplyOn[5] := TRUE;
GVL_Gr00IO.arbinGr00DoorsClosed[1] := TRUE;
GVL_Gr00IO.arbinGr00DoorsClosed[2] := TRUE;
GVL_Gr00IO.arbinGr00DoorsClosed[3] := TRUE;
GVL_Gr00IO.arbinGr00DoorsClosed[4] := TRUE;
GVL_Gr00IO.arbinGr00DoorsClosed[5] := TRUE;
GVL_Gr00IO.binGr00AllDoorsClosed := GVL_Gr00IO.arbinGr00DoorsClosed[1]
								AND GVL_Gr00IO.arbinGr00DoorsClosed[2]
								AND GVL_Gr00IO.arbinGr00DoorsClosed[3]
								AND GVL_Gr00IO.arbinGr00DoorsClosed[4]
								AND GVL_Gr00IO.arbinGr00DoorsClosed[5];

GVL_Gr00IO.binGr00AllDoorsLocked := TRUE;
GVL_Gr00IO.binGr00TempOK := TRUE;


// only for simulation
// GVL_Gr00IO.binNoEmergencyStop := TRUE;
// GVL_Gr00IO.binMoveRelease := TRUE;
// GVL_Gr00IO.binMoveReleaseSB := TRUE;
END_ACTION

END_PROGRAM

// ---- POUs/Machine/Group_0500 - Transport/Gr05MachineMode/Gr05MachineMode.TcPOU
PROGRAM Gr05MachineMode
VAR_INPUT
	(* Input variables / Eingang Variablen *)
	bEnable					:BOOL;						(* Enable Gr05MachineMode *)
END_VAR
VAR
	(* Enummerations *)

	(* Variables *)

	(* References *)

	(* Interfaces *)

	(* Instances *)

END_VAR

IF NOT bEnable
THEN
	RETURN;
END_IF;

